(* IEC 61131-3 sources: JingjiangArm/moonboxpro_arm_8.4/Application/Application/任务列表/ExtTask/动作处理/全自动套印2, 17 files *)

(* ---- EnumAutoMaticRegisterCtlMsg.st ---- *)
(*@CES
Name=EnumAutoMaticRegisterCtlMsg
Type=Gvl
TypeGuid=2db5746d-d284-4425-9f7f-2663a34b0ebc
Guid=e7e8891f-fe97-4a56-9291-de397fe1a69c
HasDeclaration=True
HasImplementation=False
*)
{DECLARATION}
// {attribute 'qualified_only'}
// {attribute 'strict'}
TYPE EnumAutoMaticRegisterCtlMsg :
(
	AMRC_MSG_NORMAL := 0,                (* 正常 *)
    AMRC_MSG_ERR_BUSY_HOR,               (* 横向正忙 *)
    AMRC_MSG_ERR_LASTAXISID_INVALID,     (* 最后一个轴id非法 *)
    AMRC_MSG_ERR_AUTOPREGISTER_VER,      (* 自动纵向套印失败 *)
    AMRC_MSG_TIMEOUT_HOR,                (* 横向预套准启动超时状态 *)
    AMRC_MSG_TIMEOUT_WAITPOS_3RD,        (* 第三方设备位置等待超时 *)
    AMRC_MSG_TIMEOUT_WAITPOS_MANU        (* 手动位置等待超时 *)
);
END_TYPE

{IMPLEMENTATION}

(* ---- EnumAutoPrintMasterStep.st ---- *)
(*@CES
Name=EnumAutoPrintMasterStep
Type=Gvl
TypeGuid=2db5746d-d284-4425-9f7f-2663a34b0ebc
Guid=e561adc0-0517-4418-b830-643ab1aeef13
HasDeclaration=True
HasImplementation=False
*)
{DECLARATION}
// 主控制状态机枚举
TYPE EnumAutoPrintMasterStep :
(
    APM_STEP_IDLE := 0,                  (* 1空闲 *)
    APM_STEP_TIPS,                       (* 2提示 *)
    APM_STEP_TIPS_ALARM,                 (* 3警铃提示 *)
    APM_STEP_AUTO_HOR,                   (* 4横向预对版 *)
    APM_STEP_AUTOING_HOR,                (* 5横向对版中 *)
    APM_STEP_AUTOSENSORPOS,              (* 6自动传感器位置 *)
    APM_STEP_SENSORPOSBYSYS3RD,          (* 7第三方设备获取传感器位置 *)
    APM_STEP_WAITPOSBY3RD,               (* 8等待第三方位置 *)
    APM_STEP_SENSORPOSBYMANU,            (* 9手动获取传感器位置 *)
    APM_STEP_WAITPOSBYMANU,              (* 10等待手动位置 *)
    APM_STEP_SENSOR_TO_TARGETPOS,        (* 11传感器到目标位置 *)
    APM_STEP_SENSOR_TO_TARGETPOSING,     (* 12传感器到目标位置中 *)
    APM_STEP_AUTO_VER,                   (* 13纵向全自动套印 *)
    APM_STEP_AUTOING_VER,                (* 14纵向全自动套印中 *)
    APM_STEP_AUTODNE_VER,                (* 15纵向全自动套印完成 *)
	APM_STEP_CALC_ADJUSTMENTS,             (** 16计算调整量 *)
    APM_STEP_FAST_ADJUSTMENT,              (** 17快速对版调整 *)
    APM_STEP_COMPLETE,                     (** 18完成 *)
    APM_STEP_TIMEOUT,                    (* 19超时 *)
    APM_STEP_ERR                         (* 20错误 *)
);
END_TYPE

{IMPLEMENTATION}

(* ---- EnumFindCommand.st ---- *)
(*@CES
Name=EnumFindCommand
Type=Gvl
TypeGuid=2db5746d-d284-4425-9f7f-2663a34b0ebc
Guid=4d4922df-cbf7-48ea-9894-b69efa7c7e4f
HasDeclaration=True
HasImplementation=False
*)
{DECLARATION}
// {attribute 'qualified_only'}
// {attribute 'strict'}
TYPE EnumFindCommand :
(
    FIND_CMD_IDLE := 0,                    (* 空闲 *)
    FIND_CMD_START_SINGLE,                 (* 开始单色寻找 *)
    FIND_CMD_START_MIX,                    (* 开始混色寻找 *)
    FIND_CMD_RESET                         (* 重置 *)
);
END_TYPE
{IMPLEMENTATION}

(* ---- EnumFindErrorCode.st ---- *)
(*@CES
Name=EnumFindErrorCode
Type=Gvl
TypeGuid=2db5746d-d284-4425-9f7f-2663a34b0ebc
Guid=764d2f18-3722-49fd-bd0f-02e1ffafaf8d
HasDeclaration=True
HasImplementation=False
*)
{DECLARATION}
// 寻找错误代码枚举
TYPE EnumFindErrorCode :
(
   	FIND_ERR_NONE := 0,                  (* 无错误 *)
    FIND_ERR_COARSE_NOT_READY := 88,     (* 粗调未到位 *)
    FIND_ERR_WAITING_CIRCLE := 50,       (* 等待1.5圈中 *)
    FIND_ERR_WAITING_FIBER_IDLE := 51,   (* 等待光纤空闲 *)
    FIND_ERR_SINGLE_MARK_NOT_FOUND := 101,(* 单色标记未找到 *)
    FIND_ERR_CALC_BEST_FAILED := 102,    (* 最佳位置计算失败 *)
    FIND_ERR_PRE_POS_INVALID := 103,     (* 前色位置无效 *)
    FIND_ERR_WAITING_SINGLE_INFO := 53,  (* 等待单色新的一圈信息 *)
    FIND_ERR_WAITING_MIX_INFO := 54,     (* 等待前色信息 *)
    FIND_ERR_TIMEOUT := 200,             (* 超时 *)
    FIND_ERR_AXIS_ID_INVALID := 201,     (* 轴ID无效 *)
    FIND_ERR_NOT_ENABLED := 202,         (* 未使能 *)
    FIND_ERR_UNKNOWN := 255              (* 未知错误 *)
);
END_TYPE
{IMPLEMENTATION}

(* ---- EnumFindState.st ---- *)
(*@CES
Name=EnumFindState
Type=Gvl
TypeGuid=2db5746d-d284-4425-9f7f-2663a34b0ebc
Guid=4b638ac6-7ee9-4b1b-9b99-b2600605b011
HasDeclaration=True
HasImplementation=False
*)
{DECLARATION}
// {attribute 'qualified_only'}
// {attribute 'strict'}
// 寻找模块状态
TYPE EnumFindState :
(
    FIND_STATE_IDLE := 0,                (* 0空闲 *)
    FIND_STATE_INIT,                     (* 1初始化 *)
    FIND_STATE_WAIT_PRESS,               (* 2等待合压 *)
    FIND_STATE_CHECK_COARSE,             (* 3检查粗调 *)
    FIND_STATE_DELAY_SINGLE,             (* 4单色前延时 *)
    FIND_STATE_FIND_SINGLE,              (* 5寻找单色 *)
    FIND_STATE_MOVE_FIBER,               (* 6移动光纤 *)
    FIND_STATE_WAIT_FIBER_MOVE,          (* 7等待光纤移动 *)
    FIND_STATE_CALC_BEST,                (* 8计算最佳位置 *)
    FIND_STATE_ADJUST_GATE,              (* 9调整波门 *)
    FIND_STATE_DELAY_MIX,                (* 10混色前延时 *)
    FIND_STATE_FINE_ADJUST,              (* 11光纤精调 *)
    FIND_STATE_WAIT_FINE_ADJ,            (* 12等待精调完成 *)
    FIND_STATE_FIND_MIX,                 (* 13寻找混色 *)
    FIND_STATE_COMPLETE,                 (* 14完成 *)
    FIND_STATE_ERROR                     (* 15错误 *)
);
END_TYPE
{IMPLEMENTATION}

(* ---- StFindResult.st ---- *)
(*@CES
Name=StFindResult
Type=Gvl
TypeGuid=2db5746d-d284-4425-9f7f-2663a34b0ebc
Guid=f624abef-a881-46ee-91b9-f19468406fe9
HasDeclaration=True
HasImplementation=False
*)
{DECLARATION}
{attribute 'pack_mode' := '1'}
// 寻找模块结果
TYPE StFindResult :
STRUCT
    xSuccess: BOOL;                      (* 寻找成功 *)
    iCurLabelPos: INT;                   (* 当前色位置 *)
    iPreLabelPos: INT;                   (* 前色位置 *)
    iCurBestPos: INT;                    (* 当前色最佳位置 *)
    rFiberMoveDist: REAL;                (* 光纤移动距离 *)
    iErrorCode: INT;                     (* 错误代码 *)
	eState: EnumFindState;				(*轴状态*)
    //sErrorMessage: STRING(255);          (* 错误信息 *)
END_STRUCT
END_TYPE
{IMPLEMENTATION}

(* ---- KS_CalBestFiberMoveDisByPS.st ---- *)
(*@CES
Name=KS_CalBestFiberMoveDisByPS
Type=FunctionBlock
TypeGuid=6f9dac99-8de1-4efc-8465-68ac443b7d08
Guid=54f61bec-2d54-4cc2-8835-56cc55fddebe
HasDeclaration=True
HasImplementation=True
*)
{DECLARATION}
FUNCTION KS_CalBestFiberMoveDisByPS : REAL
VAR_INPUT
	i_rwidth      		:POINTER TO REAL;    (*色标宽度*)
	rmark_width      : BYTE;                 (*三角形标宽度*)
    rmark_height     : BYTE;                 (*三角形标高度*)
	i_iMarkId        : INT; (*三角形标类型*)
	i_pBestMoveDisPS: POINTER TO REAL;
END_VAR
VAR
	rstandard_value  : REAL;                 (*标准宽度*)
	rdiff            : REAL;                 (*差值*)
    rdeviation       : REAL;                 (*差值乘比例*)
	rratio           : REAL;                 (*宽高比例*)
	rmove            : REAL;

END_VAR

{IMPLEMENTATION}
// 1. 安全检查：避免除零
IF (rmark_height < 1) THEN
    i_pBestMoveDisPS^ := REAL#-0.0;
    RETURN;
END_IF;

// 1. 安全检查：避免除零
IF (i_rwidth^ = 0) THEN
    i_pBestMoveDisPS^ := REAL#-0.0;
    RETURN;
END_IF;

rstandard_value := BYTE_TO_REAL(rmark_height) / 2.0;
rdiff := i_rwidth^ - rstandard_value;
rratio := BYTE_TO_REAL(rmark_width) / BYTE_TO_REAL(rmark_height);
rmove := rdiff * rratio;

// 4. 根据MARK类型决定方向
IF i_iMarkId = MARK_TYPE_TRAPE_VFLN OR i_iMarkId = MARK_TPYE_TRAPE_VBLN THEN
    i_pBestMoveDisPS^ := -rmove;  // 宽了向左调
ELSIF i_iMarkId = MARK_TYPE_TRAPE_VFLP OR i_iMarkId = MARK_TYPE_TRAPE_VBLP THEN
    i_pBestMoveDisPS^ := rmove;   // 窄了向右调
ELSIF i_iMarkId = MARK_TYPE_LINE THEN (*条标*)
	i_pBestMoveDisPS^ := 0;
END_IF;

(* ---- KS_CalBestFiberMoveDisByRS.st ---- *)
(*@CES
Name=KS_CalBestFiberMoveDisByRS
Type=FunctionBlock
TypeGuid=6f9dac99-8de1-4efc-8465-68ac443b7d08
Guid=ef5f33da-28ef-4533-8c0f-8778b1cdea74
HasDeclaration=True
HasImplementation=True
*)
{DECLARATION}
FUNCTION KS_CalBestFiberMoveDisByRS : REAL
VAR_INPUT
	i_ar_width       : ARRAY[1..3] OF REAL;    (*三个位置的色标宽度*)
	i_ar_markerpos   : ARRAY[1..3] OF INT;     (*三个色标位置信息*)
	rmark_width      : BYTE;                 (*三角形标宽度*)
    rmark_height     : BYTE;                 (*三角形标高度*)
	i_iMarkId        : INT; (*三角形标类型*)
	i_pBestPositionRS : POINTER TO INT;
	i_pBestMoveDisRS: POINTER TO REAL;
END_VAR
VAR
	i_ar_position : ARRAY[1..3] OF REAL := [0.0,-3.0,3.0];
	rstandard_value  : REAL;                 (*标准宽度*)
    ibest_index      : INT := -1;            // 最佳点索引
    rmin_diff        : REAL := REAL#1.0E6;   // 最小差值（初始值）
    iN              : INT;                   // 循环计数器
    rcurrent_diff    : REAL;                  // 当前循环计算的差值
    rbest_width      : REAL;                  // 最佳点对应的宽度
    rbest_pos        : REAL;                  // 最佳点对应的位置
    rcurrent_pos     : REAL;                  // 当前机械位置
    rwidth_ratio     : REAL;                  // 宽高比
    rdeviation       : REAL;                  // 计算出的偏差量
    rtarget_pos      : REAL;                  // 最终目标位置

END_VAR

{IMPLEMENTATION}
// 1. 安全检查：避免除零
IF (rmark_height < 1) THEN
    i_pBestMoveDisRS^ := REAL#-3.0;
    RETURN;
END_IF;

// 2. 遍历筛选最佳点（宽度最接近标准值）
ibest_index := -1;
rmin_diff := REAL#1.0E6;
rstandard_value := BYTE_TO_REAL(rmark_height) / 2;

FOR iN := 1 TO 3 DO
    // 假设位置为 -1.0 或者宽度为 -0.0 表示该点无效
    IF (i_ar_markerpos[iN] = -1 OR i_ar_width[iN] = REAL#0.0) THEN
		CONTINUE;
	ELSE
        rcurrent_diff := ABS(i_ar_width[iN] - rstandard_value);
        // 更新最佳点
        IF (rcurrent_diff < rmin_diff) THEN
            rmin_diff := rcurrent_diff;
            ibest_index := iN;
        END_IF;
    END_IF;
END_FOR;

// 3. 若无有效点，退回原点
IF (ibest_index < 0) THEN
    i_pBestMoveDisRS^ := REAL#-3.0;
    RETURN;
END_IF;

// 4. 提取计算所需数据
rbest_width := i_ar_width[ibest_index];
rbest_pos := i_ar_position[ibest_index];
rcurrent_pos := i_ar_position[3]; // 当前位置锁定为第三个点 (Index 2)

// 5. 计算几何偏差
rwidth_ratio := BYTE_TO_REAL(rmark_width) / BYTE_TO_REAL(rmark_height);
rdeviation := rmin_diff * rwidth_ratio;

// 6. 确定目标位置   以后可以改成根据色标形式控制左右方向   总体而言，是宽了往窄的方向移动，窄了往宽的方向移动
IF (i_iMarkId = MARK_TYPE_TRAPE_VFLN OR i_iMarkId = MARK_TPYE_TRAPE_VBLN) THEN
	IF (rbest_width > rstandard_value) THEN
		rtarget_pos := rbest_pos - rdeviation; // 太宽 -> 向左
	ELSIF (rbest_width < rstandard_value) THEN
		rtarget_pos := rbest_pos + rdeviation; // 太窄 -> 向右
	ELSE
		rtarget_pos := rbest_pos; // 正好
	END_IF;
ELSIF (i_iMarkId = MARK_TYPE_TRAPE_VFLP OR i_iMarkId = MARK_TYPE_TRAPE_VBLP) THEN
	IF (rbest_width > rstandard_value) THEN
		rtarget_pos := rbest_pos + rdeviation; // 太宽 -> 向右
	ELSIF (rbest_width < rstandard_value) THEN
		rtarget_pos := rbest_pos - rdeviation; // 太窄 -> 向左
	ELSE
		rtarget_pos := rbest_pos; // 正好
	END_IF;
ELSIF i_iMarkId = MARK_TYPE_LINE THEN (*条标*)
	FOR iN := 1 TO 3 DO
		// 假设位置为 -1.0 或者宽度为 -1.0 表示该点无效
		IF (i_ar_markerpos[iN] = -1 OR i_ar_width[iN] = REAL#-1.0) THEN
			CONTINUE;
		ELSE
			ibest_index := iN;
			EXIT;
		END_IF;
	END_FOR;
	(*这样可以回到零位*)
	rtarget_pos:= 0;
END_IF

// 7. 计算并返回最终移动距离
i_pBestMoveDisRS^ := rtarget_pos - rcurrent_pos;
i_pBestPositionRS^ := i_ar_markerpos[ibest_index];

(* ---- KS_CalculateMixFindDelayTime.st ---- *)
(*@CES
Name=KS_CalculateMixFindDelayTime
Type=FunctionBlock
TypeGuid=6f9dac99-8de1-4efc-8465-68ac443b7d08
Guid=2d7bebb1-5781-4f9d-9266-922f12b4caec
HasDeclaration=True
HasImplementation=True
*)
{DECLARATION}
FUNCTION KS_CalculateMixFindDelayTime  : uint
VAR_INPUT
    i_iAxisId: INT;                        (* 轴号 *)
    i_iBeforeAxisId: INT;                  (* 前轴号 *)
    i_pstUnitParam_Save: POINTER TO StUnitParam_Save; (* 单元参数 *)
    i_rVel: REAL;                          (* 速度 *)
END_VAR
VAR
    uiDelayTime: UINT;                     (* 延时时间@ms *)
    pstUnitParam_Save: POINTER TO StUnitParam_Save;
    rWaitTime: REAL;                       (* 等待时间@s *)
    rFilmLength: REAL;                     (* 料长@m *)
END_VAR
{IMPLEMENTATION}
pstUnitParam_Save := i_pstUnitParam_Save;
uiDelayTime := 0;

(* 计算前一色到此色的料长 *)
IF i_iBeforeAxisId <> -1 THEN
    (* 获取前一色到此色的料长 *)
    rFilmLength := (pstUnitParam_Save^.rFilmLengthFromPrevPressUnit)/1000.0*(i_iAxisId-i_iBeforeAxisId);

    (* 计算等待时间：料长(m) / 速度(m/min) * 60s/min = 等待时间(s) *)
    IF i_rVel > 0 THEN
        rWaitTime := rFilmLength / i_rVel * 60.0;

        (* 转换为毫秒 *)
        uiDelayTime := REAL_TO_UINT(rWaitTime * 1000.0);
    ELSE
        (* 速度为零，使用默认值 *)
        uiDelayTime := 30000;  (* 30秒 *)
    END_IF
END_IF

(* 增加安全余量（5个版周长的时间） *)
IF pstUnitParam_Save^.rGirth_PrnRoller > 0 AND i_rVel > 0 THEN
    rWaitTime := 5.0 * pstUnitParam_Save^.rGirth_PrnRoller / 1000.0 / i_rVel * 60.0;
    uiDelayTime := uiDelayTime + REAL_TO_UINT(rWaitTime * 1000.0);
END_IF

(* 最小延时时间 *)
IF uiDelayTime < 1000 THEN
    uiDelayTime := 1000;  (* 至少1秒 *)
END_IF

KS_CalculateMixFindDelayTime := uiDelayTime;

(* ---- KS_CalculateVerticalAdjustment.st ---- *)
(*@CES
Name=KS_CalculateVerticalAdjustment
Type=FunctionBlock
TypeGuid=6f9dac99-8de1-4efc-8465-68ac443b7d08
Guid=55283c42-1c2e-4d65-8dd3-8f793fe68a41
HasDeclaration=True
HasImplementation=True
*)
{DECLARATION}
(*返回计算误差的点数*)
FUNCTION KS_CalculateVerticalAdjustment : real
VAR_INPUT
    i_iAxisId: INT;                        (* 轴号 *)
    i_iCurBestSignalPos: INT;              (* 当前色最佳位置 *)
    i_iPreLabelPos: INT;                   (* 前色位置 *)
    i_pstUnitParam_Save: POINTER TO StUnitParam_Save; (* 单元参数 *)
    i_pstGrpParam_Save: POINTER TO StGrpParam_Save;  (* 组参数 *)
END_VAR
VAR
   	rAdjValue: REAL;                       (* 调整量@粗采样点数*)
    pstUnitParam_Save: POINTER TO StUnitParam_Save;
    pstGrpParam_Save: POINTER TO StGrpParam_Save;
    rTmp: REAL;
END_VAR
{IMPLEMENTATION}
pstUnitParam_Save := i_pstUnitParam_Save;
pstGrpParam_Save := i_pstGrpParam_Save;

(* 初始化返回值 *)
rAdjValue := 0.0;

(* 检查输入有效性 *)
IF i_iCurBestSignalPos >= 0 AND i_iPreLabelPos >= 0 AND
   i_iCurBestSignalPos < 4000 AND i_iPreLabelPos < 4000 THEN

    (* 根据标记排列方式计算调整量 *)
    IF pstUnitParam_Save^.iMarkArrangeMode = MARK_ARRANGE_VFOR THEN
        (* 正向排列 *)
        rTmp := INT_TO_REAL(i_iCurBestSignalPos - i_iPreLabelPos -
                   LREAL_TO_INT(20.0 * MAX_ROUNDSAMPLE_NUM / pstUnitParam_Save^.rGirth_PrnRoller));
    ELSIF pstUnitParam_Save^.iMarkArrangeMode = MARK_ARRANGE_VREV THEN
        (* 反向排列 *)
        rTmp := INT_TO_REAL(i_iCurBestSignalPos - i_iPreLabelPos +
                   LREAL_TO_INT(20.0 * MAX_ROUNDSAMPLE_NUM / pstUnitParam_Save^.rGirth_PrnRoller));
    ELSE
        (* 默认处理 *)
        rTmp := INT_TO_REAL(i_iCurBestSignalPos - i_iPreLabelPos);
    END_IF

    (* 将调整的粗采样点数转换到±MAX_ROUNDSAMPLE_NUM/2范围内 *)
    WHILE rTmp < -MAX_ROUNDSAMPLE_NUM / 2.0 DO
        rTmp := rTmp + MAX_ROUNDSAMPLE_NUM;
    END_WHILE
    WHILE rTmp > MAX_ROUNDSAMPLE_NUM / 2.0 DO
        rTmp := rTmp - MAX_ROUNDSAMPLE_NUM;
    END_WHILE

    (* 计算um单位：调整量(um) = 点数 * 版辊周长(um) / 总采样点数 *)
   // rAdjValue := rTmp * pstUnitParam_Save^.rGirth_PrnRoller * 1000.0 / MAX_ROUNDSAMPLE_NUM;
END_IF

KS_CalculateVerticalAdjustment := rTmp;

(* ---- KS_CheckSensorMotorIdleSts.st ---- *)
(*@CES
Name=KS_CheckSensorMotorIdleSts
Type=FunctionBlock
TypeGuid=6f9dac99-8de1-4efc-8465-68ac443b7d08
Guid=e3f21590-970b-415a-a0bb-786d7afe314f
HasDeclaration=True
HasImplementation=True
*)
{DECLARATION}
FUNCTION KS_CheckSensorMotorIdleSts : BOOL
(*|=0 检查所有传感器的是否处于空闲状态@所有都空闲则输出true|有一个在运动就置位false*)
(*|=合法轴id,则返回轴状态|TRUE 是空闲,FALSE是运动*)
VAR_INPUT
	i_iAxisId:INT;(*轴号@=0 *)
	i_byAxisNum:BYTE;(*轴个数@全自动套印轴*)
	i_aiAxisList_AutoAdj:ARRAY [1..MAX_UNIT_NUM] OF int;(*轴列表*)
	i_axSensorMotorIdle:ARRAY [1..MAX_UNIT_NUM] OF BOOL;(*传感器电机空闲状态@该状态不是直接通讯上来的,需要做处理后的*)
END_VAR
VAR
	iN: INT;
	xSensorMotorIdle: BOOL;
	iAxisId: INT;
	xResult: BOOL:=TRUE;
END_VAR
{IMPLEMENTATION}
IF i_iAxisId=0 THEN
	FOR iN:=2 TO i_byAxisNum BY 1 DO
		iAxisId:=i_aiAxisList_AutoAdj[iN];
		IF iAxisId>0 AND iAxisId<=MAX_UNIT_NUM THEN
			xSensorMotorIdle:=i_axSensorMotorIdle[iAxisId];
			IF NOT xSensorMotorIdle THEN(*处于运动中*)
				xResult:=FALSE;
				EXIT;
			END_IF
		END_IF
	END_FOR
ELSE
	iAxisId:=i_iAxisId;
	IF iAxisId>0 AND iAxisId<=MAX_UNIT_NUM THEN
		xSensorMotorIdle:=i_axSensorMotorIdle[iAxisId];
		IF NOT xSensorMotorIdle THEN(*处于运动中*)
			xResult:=FALSE;
		END_IF
	END_IF
END_IF

KS_CheckSensorMotorIdleSts:=xResult;

(* ---- KS_CreateTemplate.st ---- *)
(*@CES
Name=KS_CreateTemplate
Type=FunctionBlock
TypeGuid=6f9dac99-8de1-4efc-8465-68ac443b7d08
Guid=90238752-c97b-4d95-b35e-1bfe3f1964c0
HasDeclaration=True
HasImplementation=True
*)
{DECLARATION}
//构建模版函数
FUNCTION KS_CreateTemplate : BOOL
VAR_INPUT
	i_bySignalType : byte;(*模版类型，1 北人标，2普通标 ，3科赛引导条标*)
	i_iMarkTypeId : INT;(*色标形式pstStGrpParam_Save^.iMarkTypeId*)
	i_iMarkArrangeMode :INT;(*顺逆序输入*)
	i_byColorIdCurrent						: BYTE;(*当前轴色序*)
	i_rGirth_PrnRoller        :REAL;(*版周*)
	//模版构建方法 要求条标直接输入起点mm与终点mm，三角标，先确定直角边的位置，斜边按照三角标高度的一半推
	i_paiModeMidPoint:POINTER TO ARRAY [1..4] OF INT;
	i_pabyModeRadius:POINTER TO ARRAY [1..4] OF BYTE;
	i_parModeStartmm: POINTER TO ARRAY [1..4] OF REAL;
	i_parModeEndmm:POINTER TO ARRAY [1..4] OF REAL;
	i_parSignalMsg:POINTER TO ARRAY [1..15] OF REAL;
END_VAR
VAR
	iN:INT;//循环计数
	rMaxEndTemp:REAL;//记录一下最大坐标
	arStart1UMM: ARRAY [1..4] OF REAL; //mm单位 规定顺序 旗标 id 1  圆标 id 2  引导标 id 3  三角标 id 4
	arEnd1UMM: ARRAY [1..4] OF REAL; //mm单位 规定顺序 旗标 id 1  圆标 id 2  引导标 id 3  三角标 id 4
	arStart2UMM: ARRAY [1..4] OF REAL; //mm单位 规定顺序 旗标 id 1  圆标 id 2  引导标 id 3  三角标 id 4
	arEnd2UMM:ARRAY [1..4] OF REAL; //mm单位 规定顺序 旗标 id 1  圆标 id 2  引导标 id 3  三角标 id 4
	arStartMM: ARRAY [1..4] OF REAL; //mm单位 规定顺序 旗标 id 1  圆标 id 2  引导标 id 3  三角标 id 4
	arEndMM: ARRAY [1..4] OF REAL; //mm单位 规定顺序 旗标 id 1  圆标 id 2  引导标 id 3  三角标 id 4
	arStartMMTemp: ARRAY [1..4] OF REAL; //mm单位 用来导逆序，规定顺序 旗标 id 1  圆标 id 2  引导标 id 3  三角标 id 4
	arEndMMTemp: ARRAY [1..4] OF REAL; //mm单位 用来导逆序，规定顺序 旗标 id 1  圆标 id 2  引导标 id 3  三角标 id 4
	arSignalMsg:ARRAY [1..15] OF REAL; (*1旗标高度
										2 圆标高度
										3 2色引导标高度
										4 三角标高度
										5 1色旗标终点-圆标起点
										6 2色旗标终点-圆标起点
										7 1色圆标终点-引导标起点
										8 2色圆标终点-引导标起点
										9 1色引导标终点-三角标起点
										10 2色引导标终点-三角标起点
										11 2色引导标起点点-3色引导标起点
										12 1色引导标高度
*)

END_VAR

{IMPLEMENTATION}

IF 	i_parSignalMsg <> 0 AND i_rGirth_PrnRoller <> 0  THEN
	arSignalMsg:=i_parSignalMsg^;

	CASE i_bySignalType OF
	1:	//科赛引导标
		//先构建1色的模版
		arStart1UMM[1]:=  arSignalMsg[1] /2.0;//旗标起点定义旗标高度一半
		arEnd1UMM[1]:= arSignalMsg[1];//旗标终点定义旗标终点
		arStart1UMM[2]:= arEnd1UMM[1] + arSignalMsg[5];//圆标起点为旗标终点+1u5
		arEnd1UMM[2]:= arStart1UMM[2] + arSignalMsg[2];
		arStart1UMM[3]:= arEnd1UMM[2] + arSignalMsg[7];
		arEnd1UMM[3]:= arStart1UMM[3] + arSignalMsg[12];
		//条标
		IF i_iMarkTypeId = MARK_TYPE_LINE THEN
			arStart1UMM[4]:= arEnd1UMM[3] + arSignalMsg[9];
			arEnd1UMM[4]:= arStart1UMM[4] + arSignalMsg[4];
		//直角边在前
		ELSIF i_iMarkTypeId = MARK_TYPE_TRAPE_VFLP OR  i_iMarkTypeId = MARK_TYPE_TRAPE_VFLN THEN
			arStart1UMM[4]:= arEnd1UMM[3] + arSignalMsg[9];
			arEnd1UMM[4]:= arStart1UMM[4] + arSignalMsg[4]/2.0;
		ELSIF  i_iMarkTypeId = MARK_TYPE_TRAPE_VBLP OR  i_iMarkTypeId = MARK_TPYE_TRAPE_VBLN THEN
		//直角边在后
			arStart1UMM[4]:= arEnd1UMM[3] + arSignalMsg[9]+arSignalMsg[4]/2.0;
			arEnd1UMM[4]:=  arEnd1UMM[3] + arSignalMsg[9]+arSignalMsg[4];
		END_IF
		//构建2色的模版
		arStart2UMM[1]:=  arSignalMsg[1] /2.0;//旗标起点定义旗标高度一半
		arEnd2UMM[1]:= arSignalMsg[1];//旗标终点定义旗标终点
		arStart2UMM[2]:= arEnd2UMM[1] + arSignalMsg[6];
		arEnd2UMM[2]:= arStart2UMM[2] + arSignalMsg[2];
		arStart2UMM[3]:= arEnd2UMM[2] + arSignalMsg[8];
		arEnd2UMM[3]:= arStart2UMM[3] + arSignalMsg[3];
		//条标
		IF i_iMarkTypeId = MARK_TYPE_LINE THEN
			arStart2UMM[4]:= arEnd1UMM[3] + arSignalMsg[10];
			arEnd2UMM[4]:= arEnd1UMM[3] + arSignalMsg[10]+(arSignalMsg[4]);
		ELSIF i_iMarkTypeId = MARK_TYPE_TRAPE_VFLP OR  i_iMarkTypeId = MARK_TYPE_TRAPE_VFLN THEN
			arStart2UMM[4]:= arEnd1UMM[3] + arSignalMsg[10];
			arEnd2UMM[4]:= arEnd1UMM[3] + arSignalMsg[10]+(arSignalMsg[4]/2.0);
		ELSIF i_iMarkTypeId = MARK_TYPE_TRAPE_VBLP OR i_iMarkTypeId = MARK_TPYE_TRAPE_VBLN THEN
		//直角边在后
			arStart2UMM[4]:= arEnd1UMM[3] + arSignalMsg[10]+arSignalMsg[4]/2.0;
			arEnd2UMM[4]:=  arEnd1UMM[3] + arSignalMsg[10]+arSignalMsg[4];
		END_IF
		IF i_byColorIdCurrent > 0 THEN
			//根据色序选择模版
			CASE i_byColorIdCurrent OF
				1:
					FOR iN := 1 TO 4 BY 1 DO
						arStartMM[iN]:=arStart1UMM[iN];
						arEndMM[iN]:=arEnd1UMM[iN];
					END_FOR
				2:
					FOR iN := 1 TO 4 BY 1 DO
						arStartMM[iN]:=arStart2UMM[iN];
						arEndMM[iN]:=arEnd2UMM[iN];
					END_FOR
				ELSE
					arStartMM[1]:=arStart1UMM[1];
					arEndMM[1]:=arEnd1UMM[1];
					arStartMM[2]:=arStart1UMM[2]+(i_byColorIdCurrent-1)*(arSignalMsg[6]-arSignalMsg[5]);
					arEndMM[2]:=arEnd1UMM[2]+(i_byColorIdCurrent-1)*(arSignalMsg[6]-arSignalMsg[5]);
					arStartMM[3]:=arStart1UMM[3]+(i_byColorIdCurrent-1)*(arStart2UMM[3]-arStart1UMM[3]);
					arEndMM[3]:=arEnd1UMM[3]+(i_byColorIdCurrent-1)*(arEnd2UMM[3]-arEnd1UMM[3]);
					arStartMM[4]:=arStart1UMM[4]+(i_byColorIdCurrent-1)*(arStart2UMM[4]-arStart1UMM[4]);
					arEndMM[4]:=arEnd1UMM[4]+(i_byColorIdCurrent-1)*(arEnd2UMM[4]-arEnd1UMM[4]);
			END_CASE
		ELSE
			FOR iN := 1 TO 4 BY 1 DO
				arStartMM[iN]:=0;
				arEndMM[iN]:=0;
			END_FOR
		END_IF
	2: //普通标
		//关于建立没有引导,只有旗标，圆标，三角标，标建立模版，要求 3,7,8,11,12均为0，9,10填写圆标到三角标的距离，模版建立方法，虚拟一个引导标，将引导标的起点和终点与三角标相同
		//先构建1色的模版
		arStart1UMM[1]:=  arSignalMsg[1] /2.0;//旗标起点定义旗标高度一半
		arEnd1UMM[1]:= arSignalMsg[1];//旗标终点定义旗标终点
		arStart1UMM[2]:= arEnd1UMM[1] + arSignalMsg[5];//圆标起点为旗标终点+1u5
		arEnd1UMM[2]:= arStart1UMM[2] + arSignalMsg[2];

		//条标
		IF i_iMarkTypeId = MARK_TYPE_LINE THEN
			arStart1UMM[4]:= arEnd1UMM[2] + arSignalMsg[9];
			arEnd1UMM[4]:= arStart1UMM[4] + arSignalMsg[4];
			arStart1UMM[3]:= arStart1UMM[4];
			arEnd1UMM[3]:= arEnd1UMM[4];
		//直角边在前
		ELSIF i_iMarkTypeId = MARK_TYPE_TRAPE_VFLP OR  i_iMarkTypeId = MARK_TYPE_TRAPE_VFLN THEN
			arStart1UMM[4]:= arEnd1UMM[2] + arSignalMsg[9];
			arEnd1UMM[4]:= arStart1UMM[4] + arSignalMsg[4]/2.0;
			arStart1UMM[3]:= arStart1UMM[4];
			arEnd1UMM[3]:= arEnd1UMM[4];
		ELSIF  i_iMarkTypeId = MARK_TYPE_TRAPE_VBLP OR  i_iMarkTypeId = MARK_TPYE_TRAPE_VBLN THEN
		//直角边在后
			arStart1UMM[4]:= arEnd1UMM[2] + arSignalMsg[9]+arSignalMsg[4]/2.0;
			arEnd1UMM[4]:=  arEnd1UMM[2] + arSignalMsg[9]+arSignalMsg[4];
			arStart1UMM[3]:= arStart1UMM[4];
			arEnd1UMM[3]:= arEnd1UMM[4];
		END_IF
		//构建2色的模版
		arStart2UMM[1]:=  arSignalMsg[1] /2.0;//旗标起点定义旗标高度一半
		arEnd2UMM[1]:= arSignalMsg[1];//旗标终点定义旗标终点
		arStart2UMM[2]:= arEnd2UMM[1] + arSignalMsg[6];
		arEnd2UMM[2]:= arStart2UMM[2] + arSignalMsg[2];
		//条标
		IF i_iMarkTypeId = MARK_TYPE_LINE THEN
			arStart2UMM[4]:= arEnd2UMM[2] + arSignalMsg[10];
			arEnd2UMM[4]:= arStart2UMM[4] + arSignalMsg[4];
			arStart2UMM[3]:=arStart2UMM[4];
			arEnd2UMM[3]:= arEnd2UMM[4];
		//直角边在前
		ELSIF i_iMarkTypeId = MARK_TYPE_TRAPE_VFLP OR  i_iMarkTypeId = MARK_TYPE_TRAPE_VFLN THEN
			arStart2UMM[4]:= arEnd2UMM[2] + arSignalMsg[10];
			arEnd2UMM[4]:= arStart2UMM[4] + arSignalMsg[4]/2.0;
			arStart2UMM[3]:=arStart2UMM[4];
			arEnd2UMM[3]:= arEnd2UMM[4];
		ELSIF i_iMarkTypeId = MARK_TYPE_TRAPE_VBLP OR i_iMarkTypeId = MARK_TPYE_TRAPE_VBLN THEN
		//直角边在后
			arStart2UMM[4]:= arEnd2UMM[2] + arSignalMsg[10]+arSignalMsg[4]/2.0;
			arEnd2UMM[4]:=  arEnd2UMM[2] + arSignalMsg[10]+arSignalMsg[4];
			arStart2UMM[3]:=arStart2UMM[4];
			arEnd2UMM[3]:= arEnd2UMM[4];
		END_IF
		IF i_byColorIdCurrent > 0 THEN
			//根据色序选择模版
			CASE i_byColorIdCurrent OF
				1:
					FOR iN := 1 TO 4 BY 1 DO
						arStartMM[iN]:=arStart1UMM[iN];
						arEndMM[iN]:=arEnd1UMM[iN];
					END_FOR
				2:
					FOR iN := 1 TO 4 BY 1 DO
						arStartMM[iN]:=arStart2UMM[iN];
						arEndMM[iN]:=arEnd2UMM[iN];
					END_FOR
				ELSE
					arStartMM[1]:=arStart1UMM[1];
					arEndMM[1]:=arEnd1UMM[1];
					arStartMM[2]:=arStart1UMM[2]+(i_byColorIdCurrent-1)*(arSignalMsg[6]-arSignalMsg[5]);
					arEndMM[2]:=arEnd1UMM[2]+(i_byColorIdCurrent-1)*(arSignalMsg[6]-arSignalMsg[5]);
					arStartMM[4]:=arStart1UMM[4]+(i_byColorIdCurrent-1)*(arStart2UMM[4]-arStart1UMM[4]);
					arEndMM[4]:=arEnd1UMM[4]+(i_byColorIdCurrent-1)*(arEnd2UMM[4]-arEnd1UMM[4]);
					arStartMM[3]:= arStartMM[4];
					arEndMM[3]:= arEndMM[4];
			END_CASE
		ELSE
			FOR iN := 1 TO 4 BY 1 DO
				arStartMM[iN]:=0;
				arEndMM[iN]:=0;
			END_FOR
		END_IF
	3: // 3 北人标
		//先构建1色的模版
		arStart1UMM[1]:=  arSignalMsg[1] /2.0;//旗标起点定义旗标高度一半
		arEnd1UMM[1]:= arSignalMsg[1];//旗标终点定义旗标终点
		arStart1UMM[2]:= arEnd1UMM[1] + arSignalMsg[5];//圆标起点为旗标终点+1u5
		arEnd1UMM[2]:= arStart1UMM[2] + arSignalMsg[2];
		arStart1UMM[3]:= arEnd1UMM[2] + arSignalMsg[7];
		arEnd1UMM[3]:= arStart1UMM[3] + arSignalMsg[12];
		//条标
		IF i_iMarkTypeId = MARK_TYPE_LINE THEN
			arStart1UMM[4]:= arEnd1UMM[3] + arSignalMsg[9];
			arEnd1UMM[4]:= arStart1UMM[4] + arSignalMsg[4];
		//直角边在前
		ELSIF i_iMarkTypeId = MARK_TYPE_TRAPE_VFLP OR  i_iMarkTypeId = MARK_TYPE_TRAPE_VFLN THEN
			arStart1UMM[4]:= arEnd1UMM[3] + arSignalMsg[9];
			arEnd1UMM[4]:= arStart1UMM[4] + arSignalMsg[4]/2.0;
		ELSIF  i_iMarkTypeId = MARK_TYPE_TRAPE_VBLP OR  i_iMarkTypeId = MARK_TPYE_TRAPE_VBLN THEN
		//直角边在后
			arStart1UMM[4]:= arEnd1UMM[3] + arSignalMsg[9]+arSignalMsg[4]/2.0;
			arEnd1UMM[4]:=  arEnd1UMM[3] + arSignalMsg[9]+arSignalMsg[4];
		END_IF
		//构建2色的模版
		arStart2UMM[1]:=  arSignalMsg[1] /2.0;//旗标起点定义旗标高度一半
		arEnd2UMM[1]:= arSignalMsg[1];//旗标终点定义旗标终点
		arStart2UMM[2]:= arEnd2UMM[1] + arSignalMsg[6];
		arEnd2UMM[2]:= arStart2UMM[2] + arSignalMsg[2];
		arStart2UMM[3]:= arEnd2UMM[2] + arSignalMsg[8];
		arEnd2UMM[3]:= arStart2UMM[3] + arSignalMsg[3];
		//条标
		IF i_iMarkTypeId = MARK_TYPE_LINE THEN
			arStart2UMM[4]:= arEnd1UMM[3] + arSignalMsg[10];
			arEnd2UMM[4]:= arStart1UMM[4] + arSignalMsg[4];
		//直角边在前
		ELSIF i_iMarkTypeId = MARK_TYPE_TRAPE_VFLP OR  i_iMarkTypeId = MARK_TYPE_TRAPE_VFLN THEN
			arStart2UMM[4]:= arEnd2UMM[3] + arSignalMsg[10];
			arEnd2UMM[4]:= arStart2UMM[4] + arSignalMsg[4]/2.0;
		ELSIF i_iMarkTypeId = MARK_TYPE_TRAPE_VBLP OR i_iMarkTypeId = MARK_TPYE_TRAPE_VBLN THEN
		//直角边在后
			arStart2UMM[4]:= arEnd1UMM[3] + arSignalMsg[10]+arSignalMsg[4]/2.0;
			arEnd2UMM[4]:=  arEnd1UMM[3] + arSignalMsg[10]+arSignalMsg[4];
		END_IF
		IF i_byColorIdCurrent > 0 THEN
			//根据色序选择模版
			CASE i_byColorIdCurrent OF
				1:
					FOR iN := 1 TO 4 BY 1 DO
						arStartMM[iN]:=arStart1UMM[iN];
						arEndMM[iN]:=arEnd1UMM[iN];
					END_FOR
				2:
					FOR iN := 1 TO 4 BY 1 DO
						arStartMM[iN]:=arStart2UMM[iN];
						arEndMM[iN]:=arEnd2UMM[iN];
					END_FOR
				ELSE
					arStartMM[1]:=arStart1UMM[1];
					arEndMM[1]:=arEnd1UMM[1];
					arStartMM[2]:=arStart1UMM[2]+(i_byColorIdCurrent-1)*(arSignalMsg[6]-arSignalMsg[5]);
					arEndMM[2]:=arEnd1UMM[2]+(i_byColorIdCurrent-1)*(arSignalMsg[6]-arSignalMsg[5]);
					arStartMM[3]:=arStart2UMM[3]-(i_byColorIdCurrent-2)*arSignalMsg[11];
					arEndMM[3]:=arEnd2UMM[3]-(i_byColorIdCurrent-2)*arSignalMsg[11];
					arStartMM[4]:=arStart2UMM[4]+(i_byColorIdCurrent-2)*(arStart2UMM[4]-arStart1UMM[4]);
					arEndMM[4]:=arEnd2UMM[4]+(i_byColorIdCurrent-2)*(arEnd2UMM[4]-arEnd1UMM[4]);
			END_CASE
		ELSE
			FOR iN := 1 TO 4 BY 1 DO
				arStartMM[iN]:=0;
				arEndMM[iN]:=0;
			END_FOR
		END_IF
	END_CASE
	//根据顺序生成逆序模版
	IF i_iMarkArrangeMode = MARK_ARRANGE_VFOR THEN
		;//不做处理，因为本身构建是顺序的
	ELSIF i_iMarkArrangeMode = MARK_ARRANGE_VREV THEN
		FOR iN := 1 TO 4 BY 1 DO //先记录一下顺序模版
			arStartMMTemp[iN]:=arStartMM[iN];
			arEndMMTemp[iN]:=arEndMM[iN];
		END_FOR
		rMaxEndTemp:= arEndMM[4];
		FOR iN := 1 TO 4 BY 1 DO //导出逆序
			arStartMM[iN]:=rMaxEndTemp-arEndMMTemp[4-iN+1];
			arEndMM[iN]:=rMaxEndTemp-arStartMMTemp[4-iN+1];
		END_FOR
	END_IF
	FOR iN := 1 TO 4 BY 1 DO  //传出中心半径
		i_paiModeMidPoint^[iN]:=REAL_TO_INT((arEndMM[iN]+arStartMM[iN])/2.0/i_rGirth_PrnRoller*MAX_ROUNDSAMPLE_NUM);
		i_pabyModeRadius^[iN]:=REAL_TO_BYTE((arEndMM[iN]-arStartMM[iN])/2.0/i_rGirth_PrnRoller*MAX_ROUNDSAMPLE_NUM);
	END_FOR
	i_parModeStartmm^:=	arStartMM;
	i_parModeEndmm^:=arEndMM;
END_IF

(* ---- KS_FB_AutoPrintMaster.st ---- *)
(*@CES
Name=KS_FB_AutoPrintMaster
Type=FunctionBlock
TypeGuid=6f9dac99-8de1-4efc-8465-68ac443b7d08
Guid=8faa04dc-26bf-43df-9e4a-ef930424aed8
HasDeclaration=True
HasImplementation=True
*)
{DECLARATION}
FUNCTION_BLOCK KS_FB_AutoPrintMaster
VAR_INPUT
    (* 基本输入 *)
    i_xEn: BOOL;                         (* 主使能 *)
    i_rVel: REAL;                        (* 料膜速度@m/min *)
    i_rMachineryFilmLenth: REAL;         (* 机器总料长@m *)
    i_xTipsConfirm: BOOL;                (* 提示确认标志@沿触发 *)
    i_xUseAutoPreRegister_Hor: BOOL;     (* 使用横向对版功能 *)
    i_xAutoPreRegisterIdle_Hor: BOOL;    (* 横向预对版空闲状态 *)
    i_xAutoPreRegistering_Hor: BOOL;     (* 横向预对版中 *)
    i_xUseAutoSensorPos: BOOL;           (* 自动传感器位置@否则直接到纵向全自动纵向套印 *)
    i_xUseSensorPos_3rd: BOOL;           (* 使用第三方设备位置@在线|否则手动移动 *)
    i_xSensorPosValid_3rd: BOOL;         (* 传感器位置有效 *)
    i_rSenserPos_3rd: REAL;              (* 传感器位置@单位未知,暂定一个值 *)
    i_xSensorPosValid_Manu: BOOL;        (* 手动传感器值有效 *)
    i_rSensorPos_Manu: REAL;             (* 手动传感器值@绝对位置@mm *)
    i_xUseFindBestPosStep: BOOL;         (* 使用寻找最佳位置步 *)
	i_xSwitch_RFailure: BOOL;            (** R失效开关 **)
    i_xSwitch_FFailure: BOOL;            (** F失效开关 **)

    (* 轴配置 *)
    i_byAxisNum: BYTE;                   (* 轴个数@全自动套印轴 *)
    i_aiAxisList: ARRAY [1..MAX_UNIT_NUM] OF INT; (* 轴列表 *)
    i_pafbKS_FB_AxisFindModule: POINTER TO ARRAY[1..MAX_UNIT_NUM] OF KS_FB_AxisFindModule;

    (* 系统参数 *)
    i_pstStSysParam: POINTER TO StSysParam;
    i_pastStIOMap_AxisBasic: POINTER TO ARRAY [1..MAX_UNIT_NUM] OF StIOMap_Axis_FE;

    (* 快速对版参数 *)
    i_pastStAxisRapidAdjProf_V: POINTER TO ARRAY[1..MAX_UNIT_NUM] OF StAxisRapidAdjProf_V; (* 快速对版参数数组 *)

    (* 轴状态输入 *)
    i_abyRapidAdjustStep: ARRAY[1..MAX_UNIT_NUM] OF BYTE; (* 各轴快速对版步骤 *)
	i_pastFindResults :POINTER TO ARRAY[1..MAX_UNIT_NUM] OF StFindResult;
END_VAR
VAR_OUTPUT
    (* 状态输出 *)
    o_xEning: BOOL;                      (* 使能中 *)
    o_xAlarm: BOOL;                      (* 3s响铃输出 *)
   // o_xWaitingFilmLenthEn: BOOL;         (* 等料长使能 *)
    o_xAutoPreRegister_Hor: BOOL;        (* 横向自动对版@启动预套后复位 *)
   // o_xExcuteRollerPress_LastAxis: BOOL; (* 最后一个轴执行压辊动作@长有效 *)
    o_xManuConfirmSensorPos_LastAxis: BOOL; (* 最后一个轴手动确认传感器位置标志 *)

    (* 传感器电机运动 *)
    o_xSensorGoTargetPos_All: BOOL;      (* 所有轴向目标位置运动@到位后清除 *)
    o_rSenserTarPos_All: REAL;           (* 运动的目标位置 *)

    (* 动作控制 *)
    o_xExcuteAutoPreRegister_Ver: BOOL;  (* 执行纵向自动套印 *)
    o_xExcuteAutoPreRegisterDne_Ver: BOOL;(* 执行纵向自动套印完成 *)
    o_xExcuteAutoPreRegisterFailed_Ver: BOOL; (* 执行纵向自动套印失败 *)
    o_xAutoPreRegisterFinish_Ver: BOOL;  (* 执行纵向自动套印完成 *)
    o_byArcAdjAutoCtl: BYTE;             (* 套色手自动控制 *)

    (* 状态信息 *)
    o_eSts: EnumAutoPrintMasterStep;     (* 主状态机状态 *)
    o_iMsgInf: EnumAutoMaticRegisterCtlMsg; (* 信息 *)

    (* 轴控制输出 *)
    o_axAxisFindModuleEn: ARRAY[1..MAX_UNIT_NUM] OF BOOL; (* 轴寻找模块使能 *)
    o_axAxisCmd: ARRAY[1..MAX_UNIT_NUM] OF EnumFindCommand; (* 轴命令 *)

    (* 寻找结果 *)
 //   o_astFindResult: ARRAY[1..MAX_UNIT_NUM] OF StFindResult; (* 各轴寻找结果 *)
    o_xAllFindComplete: BOOL;            (* 所有轴寻找完成 *)

    (* 调整量输出 *)
    o_arAdjValue_Point: ARRAY[1..MAX_UNIT_NUM] OF REAL; (* 调整量@点 *)
    o_axAxisStartPress: ARRAY[1..MAX_UNIT_NUM] OF BOOL; (* 合压输出 *)
	o_arAdjPos_um	:ARRAY [1..MAX_UNIT_NUM] OF LREAL;(*色组调整了*)

    (* 流水线状态 *)
    o_iCurrentAxisIndex: INT;            (* 当前处理的轴索引（从后往前） *)
    o_xCurrentAxisProcessing: BOOL;      (* 当前轴正在处理 *)

    (* 轴状态显示 *)
    o_eState: ARRAY[1..MAX_UNIT_NUM] OF EnumFindState; (* 各轴状态描述 *)
	o_iErrorCode: ARRAY[1..MAX_UNIT_NUM] OF EnumFindState; (* 各轴报错*)
END_VAR
VAR
    (* 主状态机 *)
    eMainSts: EnumAutoPrintMasterStep;
    iMsgInf: EnumAutoMaticRegisterCtlMsg;

    (* 准备阶段变量 *)
    fbTimeOutTon: TON;                   (* 超时计时器 *)
    iLastAxisId: INT;                    (* 最后一个轴id *)
    rWaitFilmLenth: REAL;                (* 等待的料长@m *)
    xCheckSensorToTargetPos: BOOL;       (* 检查传感器到达目标位置 *)
    rTmp: REAL;                          (* 临时变量 *)
    xTmp: BOOL;                          (* 临时布尔 *)

    (* 传感器相关 *)
    axRollerPressSts_In: ARRAY[1..MAX_UNIT_NUM] OF BOOL; (* 压辊状态 *)
    axSensorMotorIdle: ARRAY[1..MAX_UNIT_NUM] OF BOOL;   (* 传感器电机空闲 *)

    (* 寻找结果 *)
 //   astFindResult: ARRAY[1..MAX_UNIT_NUM] OF StFindResult;

    (* 控制标志 *)
    xNextStep: BOOL;                     (* 初始化完成 *)

    (* 轴间关系 *)
    aiBeforeAxisId: ARRAY[1..MAX_UNIT_NUM] OF INT; (* 前轴号 *)
    aiAfterAxisId: ARRAY[1..MAX_UNIT_NUM] OF INT;  (* 后轴号 *)

    (* 临时变量 *)
    iN: INT;
	iM:INT;
    iAxisId: INT;
	iAxisId_Calc :INT;
    iBeforeAxisId: INT;
    iAfterAxisId: INT;

    pstStGrpParam_Save: POINTER TO StGrpParam_Save;
    pstStUnitParam_Save: POINTER TO StUnitParam_Save;
    pstStRSV_UnitParam_UnSave: POINTER TO StRSV_UnitParam_UnSave;
    pstStRSV_GrpParam_Save: POINTER TO StRSV_GrpParam_Save;

    rGirth: REAL;
    rFilmLength: REAL;

    (* 寻找结果存储 *)
    aiCurBestSignalPos: ARRAY[1..MAX_UNIT_NUM] OF INT;  (* 当前色最佳位置 *)
    aiPreLabelPos: ARRAY[1..MAX_UNIT_NUM] OF INT;       (* 前色位置 *)

    (* 轴命令控制 *)
    axAxisCmdSingle: ARRAY[1..MAX_UNIT_NUM] OF BOOL;    (* 轴单色命令触发 *)
    axAxisCmdMix: ARRAY[1..MAX_UNIT_NUM] OF BOOL;       (* 轴混色命令触发 *)

    (* 新增：简化流水线状态管理 *)
    axAxisComplete: ARRAY[1..MAX_UNIT_NUM] OF BOOL;     (* 轴完成标志 *)
    axAxisNeedPress: ARRAY[1..MAX_UNIT_NUM] OF BOOL;    (* 轴需要合压标志 *)
    axAxisPressDone: ARRAY[1..MAX_UNIT_NUM] OF BOOL;    (* 轴合压完成标志 *)
    axAxisStartPressTriggered: ARRAY[1..MAX_UNIT_NUM] OF BOOL; (* 轴合压已触发标志 *)

    (* 新增：前轴合压请求记录 *)
    axBeforeAxisPressRequested: ARRAY[1..MAX_UNIT_NUM] OF BOOL; (* 前轴合压已请求 *)

    (* 新增：所有轴完成标志 *)
    xAllAxisComplete: BOOL;               (* 所有轴完成标志 *)
	xCalculationCompleted:BOOL;           (*所有轴调整量计算完成*)

    (* 新增：轴状态描述数组 *)
  //  asAxisStatus: ARRAY[1..MAX_UNIT_NUM] OF STRING(50); (* 各轴状态描述 *)

    (* 新增：第一轴合压完成标志 *)
    xFirstAxisPressComplete: BOOL;        (* 第一轴合压完成 *)

	(*快速调整计算*)
	iIndexTmp:INT;(*//临时索引*)
	iIndex1TO2:INT;(*//从前向后的当前索引*)
	iIndex2TO1:INT;(*//从后向前的当前索引*)
	iAxisNum_1TO2:INT;(*//从前向后轴个数*)
	aiAxisIdList_FastAdj_1TO2:ARRAY [1..MAX_UNIT_NUM] OF INT;(*//从前到后压辊轴id*)
	iAxisNum_2TO1:INT;(*//从后向前轴个数*)
	aiAxisIdList_FastAdj_2TO1:ARRAY [1..MAX_UNIT_NUM] OF INT;(*//从后向前压辊轴id*)
	xCanFastAdj:BOOL;(*//可以快速对版标志*)
	iNeedFastAdjAxisNum:INT;(*//需要快速对版轴个数*)
	axFastAdjing:ARRAY [1..MAX_UNIT_NUM] OF BOOL;(*//快速对版中*)
	iAxisIdTmp:INT;
	axAdjust_ing: ARRAY [1..MAX_UNIT_NUM] OF BOOL;
	axAdjust_finish: ARRAY [1..MAX_UNIT_NUM] OF BOOL;
	xAllAdjust_finish:BOOL;
	byMeanANDAutoChangeCnt:BYTE;

END_VAR

{IMPLEMENTATION}
(* 初始化输出 *)
o_xAlarm := FALSE;
//o_xWaitingFilmLenthEn := FALSE;
o_xAutoPreRegister_Hor := FALSE;
o_xManuConfirmSensorPos_LastAxis := FALSE;
o_xSensorGoTargetPos_All := FALSE;
o_rSenserTarPos_All := 0;
o_xExcuteAutoPreRegister_Ver := FALSE;
o_xExcuteAutoPreRegisterDne_Ver := FALSE;
o_xExcuteAutoPreRegisterFailed_Ver := FALSE;
o_xAutoPreRegisterFinish_Ver := FALSE;
o_byArcAdjAutoCtl := 0;
o_xAllFindComplete := FALSE;
o_eSts := APM_STEP_IDLE;
o_iMsgInf := AMRC_MSG_NORMAL;
o_iCurrentAxisIndex := 0;
o_xCurrentAxisProcessing := FALSE;

FOR iN := 1 TO MAX_UNIT_NUM BY 1 DO
    o_axAxisFindModuleEn[iN] := FALSE;
    o_axAxisCmd[iN] := FIND_CMD_IDLE;
    i_pastFindResults^[iN].xSuccess := FALSE;
    i_pastFindResults^[iN].iErrorCode := 0;
   //
   // o_axAxisStartPress[iN] := FALSE;
  //  o_axAxisStatus[iN] := '';
END_FOR

(* 检查指针有效性 *)
IF i_pstStSysParam = 0 OR
   i_pastStIOMap_AxisBasic = 0 OR
   i_pastStAxisRapidAdjProf_V = 0 OR
   i_pafbKS_FB_AxisFindModule = 0 THEN
    RETURN;
END_IF

(* 获取外部状态 *)
FOR iN := 1 TO MAX_UNIT_NUM BY 1 DO
    pstStRSV_UnitParam_UnSave := ADR(i_pstStSysParam^.astStRSV_UnitParam_UnSave[iN]);
    axRollerPressSts_In[iN] := i_pastStIOMap_AxisBasic^[iN].o_xRel_Press;
    axSensorMotorIdle[iN] := pstStRSV_UnitParam_UnSave^.wState_FiberMove.8;
END_FOR

IF i_xEn THEN
    (* 前期准备阶段 *)
    rWaitFilmLenth := i_rMachineryFilmLenth ;  (* 等待机组料长等待 *)

    IF NOT o_xEning THEN
        (* 做参数初始化 *)
        o_xAlarm := FALSE;
        o_xAutoPreRegister_Hor := FALSE;
        o_xSensorGoTargetPos_All := FALSE;
        o_xManuConfirmSensorPos_LastAxis := FALSE;
        o_rSenserTarPos_All := 0;
        o_xExcuteAutoPreRegister_Ver := FALSE;
        o_xAutoPreRegisterFinish_Ver := FALSE;
       // o_xWaitingFilmLenthEn := FALSE;
        o_byArcAdjAutoCtl := 2;  (* 套色手动 *)

        fbTimeOutTon(IN:=FALSE);
        iLastAxisId := 0;
        xCheckSensorToTargetPos := FALSE;

        (* 计算最后一个轴ID *)
        IF i_byAxisNum > 0 AND i_byAxisNum <= MAX_UNIT_NUM THEN
            iLastAxisId := i_aiAxisList[i_byAxisNum];
        END_IF

        (* 初始化寻找结果 *)
        FOR iN := 1 TO MAX_UNIT_NUM BY 1 DO
            i_pastFindResults^[iN].xSuccess := FALSE;
            i_pastFindResults^[iN].iErrorCode := 0;
			o_arAdjValue_Point[iN] := 0.0;
			o_arAdjPos_um[iN] := 0.0;
			(* 初始化状态标志 *)
            axAxisComplete[iN] := FALSE;
            axAxisNeedPress[iN] := FALSE;
            axAxisPressDone[iN] := FALSE;
            axAxisStartPressTriggered[iN] := FALSE;
            axBeforeAxisPressRequested[iN] := FALSE;
            axAxisCmdSingle[iN] := FALSE;
            axAxisCmdMix[iN] := FALSE;
			//2026.05.19.200017+
			axAdjust_ing[iN]:=FALSE;
			axFastAdjing[iN]:=FALSE;
			axAdjust_finish[iN]:=FALSE;
        END_FOR

        (* 初始化轴间关系 *)
        FOR iN := 1 TO i_byAxisNum BY 1 DO
            iAxisId := i_aiAxisList[iN];

            (* 计算前后轴关系 *)
            IF iN = 1 THEN
                (* 第一个轴 *)
                aiBeforeAxisId[iAxisId] := -1;
                aiAfterAxisId[iAxisId] := i_aiAxisList[2];
            ELSIF iN = i_byAxisNum THEN
                (* 最后一个轴 *)
                aiBeforeAxisId[iAxisId] := i_aiAxisList[i_byAxisNum-1];
                aiAfterAxisId[iAxisId] := -1;
            ELSE
                (* 中间轴 *)
                aiBeforeAxisId[iAxisId] := i_aiAxisList[iN-1];
                aiAfterAxisId[iAxisId] := i_aiAxisList[iN+1];
            END_IF
		   //o_axAxisStartPress[iAxisId] := TRUE;
          //  asAxisStatus[iAxisId] := '空闲';
        END_FOR
		xNextStep:=TRUE;
		FOR iN:=2 TO i_byAxisNum BY 1 DO(*开始的时候全部打手动*)
			iAxisId:= i_aiAxisList[iN];
			pstStUnitParam_Save:= ADR(i_pstStsysParam^.astStUnitParam_Save[iAxisId]);
			IF pstStUnitParam_Save^.dwFlag_Sts.0 OR pstStUnitParam_Save^.dwFlag_Sts.1 THEN
				pstStUnitParam_Save^.dwFlag_Sts.0:= FALSE;
				pstStUnitParam_Save^.dwFlag_Sts.1:= FALSE;
				xNextStep:=FALSE;
			END_IF
		END_FOR
        (* 初始化全自动控制变量 *)
        xAllAxisComplete := FALSE;
        xFirstAxisPressComplete := FALSE;
		xCanFastAdj:=FALSE;

        IF xNextStep THEN
			o_xEning := TRUE;
			eMainSts := APM_STEP_TIPS;
			iMsgInf := AMRC_MSG_NORMAL;
		END_IF
      //  xInitDone := FALSE;
    END_IF

    (* 主状态机处理 - 前期准备阶段 *)
    CASE eMainSts OF
        APM_STEP_IDLE:
            (* 空闲状态 *)
            ;

        APM_STEP_TIPS:
            IF i_xTipsConfirm THEN
                eMainSts := APM_STEP_TIPS_ALARM;
            END_IF

        APM_STEP_TIPS_ALARM:
            o_xAlarm := TRUE;
            fbTimeOutTon(IN:=TRUE, PT:=T#3S);

            IF fbTimeOutTon.Q THEN
                IF i_xUseAutoPreRegister_Hor THEN
                    eMainSts := APM_STEP_AUTO_HOR;
                ELSE
                    IF i_xUseAutoSensorPos THEN
                        eMainSts := APM_STEP_AUTOSENSORPOS;
                    ELSE
                        eMainSts := APM_STEP_AUTO_VER;
                    END_IF
                END_IF
            END_IF

            (* 复位计时器 *)
            IF eMainSts <> APM_STEP_TIPS_ALARM THEN
                o_xAlarm := FALSE;
                fbTimeOutTon(IN:=FALSE);
            END_IF

        (* 横向动作状态处理 *)
        APM_STEP_AUTO_HOR:
            IF i_xAutoPreRegisterIdle_Hor THEN
                o_xAutoPreRegister_Hor := TRUE;

                IF i_xAutoPreRegistering_Hor THEN
                    eMainSts := APM_STEP_AUTOING_HOR;
                ELSE
                    fbTimeOutTon(IN:=TRUE, PT:=T#1S);
                    IF fbTimeOutTon.Q THEN
                        eMainSts := APM_STEP_TIMEOUT;
                    END_IF
                END_IF
            ELSE
                eMainSts := APM_STEP_ERR;
            END_IF

            (* 错误信息处理 *)
            IF eMainSts = APM_STEP_ERR THEN
                iMsgInf := AMRC_MSG_ERR_BUSY_HOR;
            END_IF
            IF eMainSts = APM_STEP_TIMEOUT THEN
                iMsgInf := AMRC_MSG_TIMEOUT_HOR;
            END_IF

            (* 退出case复位计时器 *)
            IF eMainSts <> APM_STEP_AUTO_HOR THEN
                o_xAutoPreRegister_Hor := FALSE;
                fbTimeOutTon(IN:=FALSE);
            END_IF

        APM_STEP_AUTOING_HOR:
            IF NOT i_xAutoPreRegistering_Hor THEN
                IF i_xUseAutoSensorPos THEN
                    eMainSts := APM_STEP_AUTOSENSORPOS;
                ELSE
                    eMainSts := APM_STEP_AUTO_VER;
                END_IF
            END_IF

        (* 自动sensor位置控制 *)
        APM_STEP_AUTOSENSORPOS:
            IF i_xUseSensorPos_3rd THEN
                eMainSts := APM_STEP_SENSORPOSBYSYS3RD;
            ELSE
                eMainSts := APM_STEP_SENSORPOSBYMANU;
            END_IF

        (* 第三方设备获取传感器位置 *)
        APM_STEP_SENSORPOSBYSYS3RD:
            IF iLastAxisId <> 0 THEN
                IF NOT axRollerPressSts_In[iLastAxisId] THEN
					o_axAxisStartPress[iLastAxisId] := TRUE;
                    //o_xExcuteRollerPress_LastAxis := TRUE;
                END_IF
                eMainSts := APM_STEP_WAITPOSBY3RD;
            ELSE
                eMainSts := APM_STEP_ERR;
            END_IF

            IF eMainSts = APM_STEP_ERR THEN
                iMsgInf := AMRC_MSG_ERR_LASTAXISID_INVALID;
            END_IF

        APM_STEP_WAITPOSBY3RD:
            IF NOT i_xSensorPosValid_3rd THEN
                eMainSts := APM_STEP_SENSOR_TO_TARGETPOS;
                o_rSenserTarPos_All := i_rSenserPos_3rd;
            ELSE
                IF i_rVel <> 0 THEN
                    rTmp := rWaitFilmLenth / i_rVel * 60;
                ELSE
                    rTmp := rWaitFilmLenth / 30.0 * 60;
                END_IF
                rTmp := rTmp * 1000;  (* 转换为毫秒 *)

                fbTimeOutTon(IN:=TRUE, PT:=REAL_TO_TIME(rTmp));
                IF fbTimeOutTon.Q THEN
                    eMainSts := APM_STEP_TIMEOUT;
                END_IF
            END_IF

            (* 输出信息 *)
            IF eMainSts = APM_STEP_TIMEOUT THEN
                iMsgInf := AMRC_MSG_TIMEOUT_WAITPOS_3RD;
            END_IF

            IF eMainSts <> APM_STEP_WAITPOSBY3RD THEN
                fbTimeOutTon(IN:=FALSE);
            END_IF

        (* 手动确认传感器位置 *)
        APM_STEP_SENSORPOSBYMANU:
            IF iLastAxisId <> 0 THEN
                IF NOT axRollerPressSts_In[iLastAxisId] THEN
					o_axAxisStartPress[iLastAxisId] := TRUE;
                    //o_xExcuteRollerPress_LastAxis := TRUE;
                END_IF
                eMainSts := APM_STEP_WAITPOSBYMANU;
            ELSE
                eMainSts := APM_STEP_ERR;
            END_IF

            IF eMainSts = APM_STEP_ERR THEN
                iMsgInf := AMRC_MSG_ERR_LASTAXISID_INVALID;
            END_IF

        APM_STEP_WAITPOSBYMANU:
            o_xManuConfirmSensorPos_LastAxis := TRUE;

            IF  i_xSensorPosValid_Manu THEN
                eMainSts := APM_STEP_SENSOR_TO_TARGETPOS;
                o_rSenserTarPos_All := i_rSensorPos_Manu;
            ELSE
                IF i_rVel <> 0 THEN
                    rTmp := rWaitFilmLenth / i_rVel * 60;
                ELSE
                    rTmp := rWaitFilmLenth / 30.0 * 60;;
                END_IF
                rTmp := rTmp * 1000;  (* 转换为毫秒 *)

                fbTimeOutTon(IN:=TRUE, PT:=REAL_TO_TIME(rTmp));
                IF fbTimeOutTon.Q THEN
                    eMainSts := APM_STEP_TIMEOUT;
                END_IF
            END_IF

            (* 输出信息 *)
            IF eMainSts = APM_STEP_TIMEOUT THEN
                iMsgInf := AMRC_MSG_TIMEOUT_WAITPOS_MANU;
            END_IF

            IF eMainSts <> APM_STEP_WAITPOSBYMANU THEN
                fbTimeOutTon(IN:=FALSE);
                o_xManuConfirmSensorPos_LastAxis := FALSE;
            END_IF

        (* 传感器电机向目标位置运动 *)
        APM_STEP_SENSOR_TO_TARGETPOS:
            xTmp := KS_CheckSensorMotorIdleSts(0, i_byAxisNum, i_aiAxisList, axSensorMotorIdle);
            IF xTmp THEN
                o_xSensorGoTargetPos_All := TRUE;
            END_IF

            IF o_xSensorGoTargetPos_All THEN
				eMainSts := APM_STEP_SENSOR_TO_TARGETPOSING;
				o_xSensorGoTargetPos_All := FALSE;
            END_IF

        APM_STEP_SENSOR_TO_TARGETPOSING:
            xTmp := KS_CheckSensorMotorIdleSts(iLastAxisId, i_byAxisNum, i_aiAxisList, axSensorMotorIdle);

            IF i_xUseFindBestPosStep THEN
                xCheckSensorToTargetPos := TRUE;
                eMainSts := APM_STEP_AUTO_VER;
            ELSE
                IF xTmp THEN
                    eMainSts := APM_STEP_AUTO_VER;
                END_IF
            END_IF

        (* 纵向全自动套印 - 流水线处理 *)
        APM_STEP_AUTO_VER:
            (* 启动寻找模块 *)
            o_xExcuteAutoPreRegister_Ver := TRUE;
            o_xCurrentAxisProcessing := TRUE;
            axAxisNeedPress[iLastAxisId]:=TRUE;
            eMainSts := APM_STEP_AUTOING_VER;

        APM_STEP_AUTOING_VER:
            (* 简化流水线处理逻辑 - 只负责触发前轴合压和激活寻找模块 *)
            o_xCurrentAxisProcessing := TRUE;
            o_iCurrentAxisIndex := 0;

            (* 首先，更新所有轴的状态描述 *)
            xAllAxisComplete := TRUE;  (* 假设所有轴都完成 *)

            FOR iN := i_byAxisNum TO 1 BY -1 DO
                iAxisId := i_aiAxisList[iN];
                iBeforeAxisId := aiBeforeAxisId[iAxisId];

                (* 跳过已完成的轴 *)
                IF axAxisComplete[iAxisId] THEN
                    CONTINUE;
                END_IF

                (* 标记有轴未完成 *)
                xAllAxisComplete := FALSE;

                (* 记录当前正在处理的轴索引 *)
                IF NOT axAxisComplete[iAxisId] THEN
                    o_iCurrentAxisIndex := iN;
                END_IF

                (* 第一轴特殊处理：只需要合压 *)
                IF iN = 1 THEN
                    (* 第一轴尚未合压完成 *)
                    IF NOT axAxisPressDone[iAxisId] THEN
                        (* 检查是否需要合压 *)
                        IF axAxisNeedPress[iAxisId] AND NOT axAxisPressDone[iAxisId] THEN
                            (* 触发合压 *)
                            IF NOT axAxisStartPressTriggered[iAxisId] THEN
                                o_axAxisStartPress[iAxisId] := TRUE;
                                axAxisStartPressTriggered[iAxisId] := TRUE;
                              //  asAxisStatus[iAxisId] := '合压中';
                            END_IF

                            (* 检查合压是否完成 *)
                            IF axRollerPressSts_In[iAxisId] THEN
                                (* 合压完成 *)
                                o_axAxisStartPress[iAxisId] := FALSE;
                                axAxisPressDone[iAxisId] := TRUE;
                                axAxisComplete[iAxisId] := TRUE;
                             //   asAxisStatus[iAxisId] := '完成';
                                xFirstAxisPressComplete := TRUE;
                            END_IF
                        END_IF
                    END_IF
                    CONTINUE;
                END_IF

                (* 非第一轴的处理逻辑 *)

                (* 1. 检查是否需要合压 *)
                IF axAxisNeedPress[iAxisId] AND NOT axAxisPressDone[iAxisId] THEN
                    (* 需要合压但未合压 *)
                    IF NOT axAxisStartPressTriggered[iAxisId] THEN
                        (* 触发合压 *)
                        IF iN = i_byAxisNum THEN
                            (* 最后一个轴 *)
							o_axAxisStartPress[iLastAxisId] := TRUE;
                        ELSE
                            (* 其他轴 *)
                            o_axAxisStartPress[iAxisId] := TRUE;
                        END_IF
                        axAxisStartPressTriggered[iAxisId] := TRUE;
                     //   asAxisStatus[iAxisId] := '等待合压';
                    END_IF

                    (* 检查合压是否完成 *)
                    IF axRollerPressSts_In[iAxisId] THEN
                        (* 合压完成 *)
//                         IF iN = i_byAxisNum THEN
// 							o_axAxisStartPress[iLastAxisId] := TRUE;
//                         END_IF
                        o_axAxisStartPress[iAxisId] := FALSE;
                        axAxisPressDone[iAxisId] := TRUE;

                        (* 激活寻找模块并发送单色寻找命令 *)
                        o_axAxisFindModuleEn[iAxisId] := TRUE;
                        IF NOT axAxisCmdSingle[iAxisId] THEN
                            o_axAxisCmd[iAxisId] := FIND_CMD_START_SINGLE;
                            axAxisCmdSingle[iAxisId] := TRUE;
                        END_IF

                      //  asAxisStatus[iAxisId] := '寻找单色中';
                    END_IF
                END_IF

                (* 2. 检查轴寻找模块的状态 *)
                IF axAxisPressDone[iAxisId] AND NOT axAxisComplete[iAxisId] THEN
                    (* 轴已合压完成，正在寻找中 *)

                    (* 激活寻找模块 *)
                    o_axAxisFindModuleEn[iAxisId] := TRUE;

                    (* 3. 检查是否需要触发前轴合压 *)
                    IF iBeforeAxisId <> -1 THEN
                        (* 检查轴寻找模块是否发出前轴合压信号 *)
                        IF i_pafbKS_FB_AxisFindModule^[iAxisId].o_xBeforeAxisStartPress AND
                           NOT axBeforeAxisPressRequested[iAxisId] THEN
                            (* 触发前轴合压 *)
                            axAxisNeedPress[iBeforeAxisId] := TRUE;
                            axBeforeAxisPressRequested[iAxisId] := TRUE;
                        END_IF
                    END_IF

                    (* 4. 检查轴是否完成 *)
                    IF i_pafbKS_FB_AxisFindModule^[iAxisId].o_xDone THEN
                        (* 轴寻找完成 *)
                        o_axAxisFindModuleEn[iAxisId] := FALSE;
                        axAxisComplete[iAxisId] := TRUE;

                        (* 保存寻找结果 *)
                        i_pastFindResults^[iAxisId] := i_pafbKS_FB_AxisFindModule^[iAxisId].o_stResult;
                        aiCurBestSignalPos[iAxisId] := i_pastFindResults^[iAxisId].iCurBestPos;

                        (* 记录前色位置（如果找到混色）*)
                        IF i_pastFindResults^[iAxisId].iPreLabelPos >= 0 THEN
                            aiPreLabelPos[iAxisId] := i_pastFindResults^[iAxisId].iPreLabelPos;
                        END_IF

                        (* 复位命令 *)
                        IF axAxisCmdSingle[iAxisId] THEN
                            o_axAxisCmd[iAxisId] := FIND_CMD_IDLE;
                            axAxisCmdSingle[iAxisId] := FALSE;
                        END_IF

                        IF axAxisCmdMix[iAxisId] THEN
                            o_axAxisCmd[iAxisId] := FIND_CMD_IDLE;
                            axAxisCmdMix[iAxisId] := FALSE;
                        END_IF
                    END_IF
                END_IF
            END_FOR

            (* 检查是否所有轴都完成 *)
            IF xAllAxisComplete THEN
                eMainSts := APM_STEP_CALC_ADJUSTMENTS;
                (* 复位全自动套印标志 *)
                o_xExcuteAutoPreRegister_Ver := FALSE;
                o_xAutoPreRegisterFinish_Ver := TRUE;
            END_IF

        APM_STEP_CALC_ADJUSTMENTS:
            (* 计算调整量 *)
           // o_xBusy := TRUE;

            (* 计算每个轴的调整量（从第二个轴开始）*)
            FOR iN := 2 TO i_byAxisNum BY 1 DO
                iAxisId := i_aiAxisList[iN];

                (* 获取参数指针 *)
                pstStUnitParam_Save := ADR(i_pstStSysParam^.astStUnitParam_Save[iAxisId]);
                pstStGrpParam_Save := ADR(i_pstStSysParam^.astStGrpParam_Save);

                (* 计算纵向调整量 *)
                IF aiCurBestSignalPos[iAxisId] >= 0 AND aiPreLabelPos[iAxisId] >= 0 THEN
                    o_arAdjValue_Point[iAxisId] := KS_CalculateVerticalAdjustment(
                        iAxisId,
                        aiCurBestSignalPos[iAxisId],
                        aiPreLabelPos[iAxisId],
                        pstStUnitParam_Save,
                        pstStGrpParam_Save
                    );
                ELSE
                    o_arAdjValue_Point[iAxisId] := 0.0;
                END_IF
            END_FOR
            xCalculationCompleted:=FALSE;
			(*动作执行*)

			FOR iN:=2 TO i_byAxisNum BY 1 DO
				iAxisId:=i_aiAxisList[iN];
				pstStUnitParam_Save:= ADR(i_pstStsysParam^.astStUnitParam_Save[iAxisId]);
				o_arAdjPos_um[iAxisId]:=0;
				FOR iM:=2 TO iN BY 1 DO
					iAxisId_Calc:= i_aiAxisList[iM];
					(*当前色获取到的粗采样点数*)
					rTmp:=o_arAdjValue_Point[iAxisId_Calc];(*记录位置*)
					(*累加@此时单位还是粗采样点数*)
					o_arAdjPos_um[iAxisId]:=o_arAdjPos_um[iAxisId] + rTmp;
				END_FOR
				(*测试*)
				//o_arAdjPos_um[iAxisId]:=15000*iAxisId;
				(*2026.3.26.213041+ by liu.yt*)
				(*将调整的粗采样点数转换到+-MAX_ROUNDSAMPLE_NUM/2范围内*)
				WHILE o_arAdjPos_um[iAxisId] < -MAX_ROUNDSAMPLE_NUM / 2 DO
					o_arAdjPos_um[iAxisId] := o_arAdjPos_um[iAxisId] + MAX_ROUNDSAMPLE_NUM;
				END_WHILE
				WHILE o_arAdjPos_um[iAxisId] > MAX_ROUNDSAMPLE_NUM / 2 DO
					o_arAdjPos_um[iAxisId] := o_arAdjPos_um[iAxisId] - MAX_ROUNDSAMPLE_NUM;
				END_WHILE(*此时单位还是粗采样点数*)
				(*计算um单位*)
				o_arAdjPos_um[iAxisId]:= o_arAdjPos_um[iAxisId]* pstStUnitParam_Save^.rGirth_PrnRoller*1000 / MAX_ROUNDSAMPLE_NUM;
			END_FOR
			xCalculationCompleted:=TRUE;
            (* 进入快速调整步骤 *)
            eMainSts := APM_STEP_FAST_ADJUSTMENT;

        APM_STEP_FAST_ADJUSTMENT:
            (* 快速对版调整 *)
            //o_xBusy := TRUE;
			Action_Excute();
			IF xAllAdjust_finish THEN
				eMainSts := APM_STEP_COMPLETE;
				byMeanANDAutoChangeCnt:=0;
			END_IF
        APM_STEP_COMPLETE:
            (* 完成 *)
           // o_xBusy := FALSE;
		   IF xAllAdjust_finish THEN(*全部调整完成-自动合压*)
			   xNextStep:=TRUE;
				FOR iN:=2 TO i_byAxisNum BY 1 DO(*开始的时候全部打手动*)
					iAxisId:= i_aiAxisList[iN];
					pstStUnitParam_Save:= ADR(i_pstStsysParam^.astStUnitParam_Save[iAxisId]);
					(*结束后全部打自动*)
					IF NOT pstStUnitParam_Save^.dwFlag_Sts.0 THEN
						pstStUnitParam_Save^.dwFlag_Sts.0:= TRUE;
						xNextStep:=FALSE;
					END_IF
				END_FOR
				IF xNextStep THEN
					o_xAllFindComplete := TRUE;
				END_IF

// 				byMeanANDAutoChangeCnt := byMeanANDAutoChangeCnt+1;
// 				IF  byMeanANDAutoChangeCnt < 3 THEN
// 					o_byArcAdjAutoCtl:=1;
// 					o_xWaitingFilmLenthEn := TRUE;
// 				ELSE
// 					o_xWaitingFilmLenthEn := FALSE;
//
// 					//xAllAdjust_finish:=FALSE;
// 				END_IF
			END_IF

        (* 超时步 *)
        APM_STEP_TIMEOUT:
            eMainSts := APM_STEP_ERR;
            iMsgInf := AMRC_MSG_TIMEOUT_HOR;

        (* 返回失败 *)
        APM_STEP_ERR:
            o_xExcuteAutoPreRegisterFailed_Ver := TRUE;
            o_xAllFindComplete := FALSE;
    END_CASE

    (* 调用所有轴的寻找模块 *)
    FOR iN := 1 TO i_byAxisNum BY 1 DO
        iAxisId := i_aiAxisList[iN];

        (* 获取参数指针 *)
        pstStRSV_UnitParam_UnSave := ADR(i_pstStSysParam^.astStRSV_UnitParam_UnSave[iAxisId]);
        pstStUnitParam_Save := ADR(i_pstStSysParam^.astStUnitParam_Save[iAxisId]);
        pstStGrpParam_Save := ADR(i_pstStSysParam^.astStGrpParam_Save);
        pstStRSV_GrpParam_Save := ADR(i_pstStSysParam^.astStRSV_GrpParam_Save);

        rGirth := pstStUnitParam_Save^.rGirth_PrnRoller;
        rFilmLength := pstStUnitParam_Save^.rFilmLengthFromPrevPressUnit;

        (* 获取前后轴号 *)
        iBeforeAxisId := aiBeforeAxisId[iAxisId];
        iAfterAxisId := aiAfterAxisId[iAxisId];

        (* 调用轴寻找模块 *)
        i_pafbKS_FB_AxisFindModule^[iAxisId](
            (* 基本输入 *)
            i_xEn := o_axAxisFindModuleEn[iAxisId],
            i_iAxisId := iAxisId,
            i_eCmd := o_axAxisCmd[iAxisId],
            i_xUseFindBestPosStep := i_xUseFindBestPosStep,

            (* 参数输入 *)
            i_pstStRSV_UnitParam_UnSave := pstStRSV_UnitParam_UnSave,
            i_pstStUnitParam_Save := pstStUnitParam_Save,
            i_pstStGrpParam_Save := pstStGrpParam_Save,
            i_rVel := i_rVel,
            i_rGirth := rGirth,
            i_rFilmLength := rFilmLength,
            i_iBeforeAxisId := iBeforeAxisId,
            i_iAfterAxisId := iAfterAxisId,
            i_rFindBestPos_MoveDis := pstStRSV_GrpParam_Save^.arFiberMove,

            (* 外部状态输入 *)
            i_xCoarseDone := axSensorMotorIdle[iAxisId],
            i_xPressDone := axRollerPressSts_In[iAxisId],
            i_xAutoMode := (eMainSts = APM_STEP_AUTOING_VER),
            i_xFind_IDLE := pstStRSV_UnitParam_UnSave^.byFlag_CommFromSlave.4,

            (* 开关参数 *)
            i_xSwitch_EnFastPress := pstStRSV_GrpParam_Save^.xSwitch_EnFastPress,
            i_xSwitch_RFailure := FALSE,
            i_xSwitch_FFailure := FALSE,
            i_xSpecialMarkEn := FALSE
        );

    END_FOR

ELSE
    (* 复位处理 *)
    IF o_xEning THEN
        o_xEning := FALSE;
        eMainSts := APM_STEP_IDLE;
        o_xAlarm := FALSE;
        o_xAutoPreRegister_Hor := FALSE;
        o_xManuConfirmSensorPos_LastAxis := FALSE;
        o_xSensorGoTargetPos_All := FALSE;
        o_rSenserTarPos_All := 0;
        o_xExcuteAutoPreRegister_Ver := FALSE;
      //  o_xWaitingFilmLenthEn := FALSE;
        xCheckSensorToTargetPos := FALSE;
        o_byArcAdjAutoCtl := 0;  (* 套色手动 *)
		xCalculationCompleted:=FALSE;
        (* 复位所有轴的寻找模块 *)
		FOR iN:=1 TO MAX_UNIT_NUM BY 1 DO
			 o_axAxisStartPress[iAxisId]:=FALSE;
		END_FOR
        FOR iN := 1 TO i_byAxisNum BY 1 DO
            iAxisId := i_aiAxisList[iN];
            (* 获取参数指针 *)
            pstStRSV_UnitParam_UnSave := ADR(i_pstStSysParam^.astStRSV_UnitParam_UnSave[iAxisId]);
            pstStUnitParam_Save := ADR(i_pstStSysParam^.astStUnitParam_Save[iAxisId]);
            pstStGrpParam_Save := ADR(i_pstStSysParam^.astStGrpParam_Save);
            pstStRSV_GrpParam_Save := ADR(i_pstStSysParam^.astStRSV_GrpParam_Save);

            rGirth := pstStUnitParam_Save^.rGirth_PrnRoller;
            rFilmLength := pstStUnitParam_Save^.rFilmLengthFromPrevPressUnit;

            (* 获取前后轴号 *)
            iBeforeAxisId := aiBeforeAxisId[iAxisId];
            iAfterAxisId := aiAfterAxisId[iAxisId];

            (* 调用轴寻找模块复位 *)
            i_pafbKS_FB_AxisFindModule^[iAxisId](
                (* 基本输入 *)
                i_xEn := TRUE,
                i_iAxisId := iAxisId,
                i_eCmd := FIND_CMD_RESET,
                i_xUseFindBestPosStep := i_xUseFindBestPosStep,

                (* 参数输入 *)
                i_pstStRSV_UnitParam_UnSave := pstStRSV_UnitParam_UnSave,
                i_pstStUnitParam_Save := pstStUnitParam_Save,
                i_pstStGrpParam_Save := pstStGrpParam_Save,
                i_rVel := i_rVel,
                i_rGirth := rGirth,
                i_rFilmLength := rFilmLength,
                i_iBeforeAxisId := iBeforeAxisId,
                i_iAfterAxisId := iAfterAxisId,
				i_rFindBestPos_MoveDis := pstStRSV_GrpParam_Save^.arFiberMove,

                (* 外部状态输入 *)
                i_xCoarseDone := pstStRSV_UnitParam_UnSave^.wState_FiberMove.8,
                i_xPressDone := axRollerPressSts_In[iAxisId],
                i_xAutoMode := FALSE,
                i_xFind_IDLE := pstStRSV_UnitParam_UnSave^.byFlag_CommFromSlave.4,

                (* 开关参数 *)
                i_xSwitch_EnFastPress := pstStRSV_GrpParam_Save^.xSwitch_EnFastPress,
                i_xSwitch_RFailure := i_xSwitch_RFailure,
                i_xSwitch_FFailure := i_xSwitch_FFailure,
                i_xSpecialMarkEn := FALSE
            );
			i_pastFindResults^[iAxisId] := i_pafbKS_FB_AxisFindModule^[iAxisId].o_stResult;
        END_FOR
    END_IF
END_IF

(* 输出状态 *)
o_eSts := eMainSts;
o_iMsgInf := iMsgInf;
//o_astFindResult := astFindResult;
g_axAutoFind_Press:=o_axAxisStartPress;
FOR iN := 1 TO i_byAxisNum BY 1 DO
	iAxisId := i_aiAxisList[iN];
	o_eState[iAxisId]:= i_pafbKS_FB_AxisFindModule^[iAxisId].o_eState;
	o_iErrorCode[iAxisId]:=i_pafbKS_FB_AxisFindModule^[iAxisId].o_stResult.iErrorCode;
END_FOR

//o_axAxisStatus := asAxisStatus;

(* ---- KS_FB_AxisFindModule.st ---- *)
(*@CES
Name=KS_FB_AxisFindModule
Type=FunctionBlock
TypeGuid=6f9dac99-8de1-4efc-8465-68ac443b7d08
Guid=fe608f45-03e0-4e2e-a249-20c440ac82a6
HasDeclaration=True
HasImplementation=True
*)
{DECLARATION}
FUNCTION_BLOCK KS_FB_AxisFindModule
VAR_INPUT
    (** 基本输入 **)
    i_xEn: BOOL;                         (** 模块使能 **)
    i_iAxisId: INT;                      (** 轴号 **)
    i_eCmd: EnumFindCommand;             (** 命令 **)
    i_xUseFindBestPosStep: BOOL;         (** 使用寻找最佳位置步骤 **)

    (** 参数输入 **)
    i_pstStRSV_UnitParam_UnSave: POINTER TO StRSV_UnitParam_UnSave; (** 单元参数 **)
    i_pstStUnitParam_Save: POINTER TO StUnitParam_Save; (** 单元参数 **)
    i_pstStGrpParam_Save: POINTER TO StGrpParam_Save; (** 组参数 **)
    i_rVel: REAL;                        (** 速度 **)
    i_rGirth: REAL;                      (** 版周长 **)
    i_rFilmLength: REAL;                 (** 料长 **)
    i_iBeforeAxisId: INT;                (** 前轴号 **)
    i_iAfterAxisId: INT;                 (** 后轴号 **)
    i_rFindBestPos_MoveDis: ARRAY [1..2] OF REAL; (** 光纤移动距离 **)

    (** 外部状态输入 **)
    i_xCoarseDone: BOOL;                 (** 粗调完成标志 **)
    i_xPressDone: BOOL;                  (** 合压完成标志 **)
    i_xAutoMode: BOOL;                   (** 自动模式标志 **)
    i_xFind_IDLE: BOOL;                  (** 当前轴全自动套印空闲 **)

    (** 开关参数 **)
    i_xSwitch_EnFastPress: BOOL;         (** 快速合压开关 **)
    i_xSwitch_RFailure: BOOL;            (** R失效开关 **)
    i_xSwitch_FFailure: BOOL;            (** F失效开关 **)
    i_xSpecialMarkEn: BOOL;              (** 特殊标使能 **)
END_VAR
VAR_OUTPUT
    (** 状态输出 **)
    o_eState: EnumFindState;             (** 当前状态 **)
    o_stResult: StFindResult;            (** 寻找结果 **)
    o_xBusy: BOOL;                       (** 忙标志 **)
    o_xDone: BOOL;                       (** 完成标志 **)
    o_xSuccess: BOOL;                    (** 成功标志 **)
    o_xError: BOOL;                      (** 错误标志 **)
    o_iErrorCode: INT;                   (** 错误代码 **)

    (** 控制输出 **)
    o_xNeedPress: BOOL;                  (** 需要合压 **)
    o_xBeforeAxisStartPress: BOOL;       (** 前轴开始合压（自动模式下使用）**)

    (** 从站控制信号 **)
    o_xFindFirstMark: BOOL;              (** 启动单色寻找@发送给从站 **)
    o_xFindPreMark: BOOL;                (** 启动混色寻找@发送给从站 **)
    o_xGateMoveFinish: BOOL;             (** 波门移动完成 **)
    o_xCurManuAdjust: BOOL;              (** 当前色需要手动调整 **)
    o_xPreCurManuAdjust: BOOL;           (** 前色需要手动调整 **)

    (** 光纤移动控制 **)
    o_xFiberMoveDisRunStart_FindSignal: BOOL; (** 光纤移动启动 **)
    o_rFiberMoveDistanceIn_FindSignal: REAL; (** 光纤移动距离 **)

    (** 参数设置输出 **)
    o_iGateSa: INT;                      (** 波门起始位置 **)

    (** 寻找状态标志 **)
    o_xSingleFound: BOOL;                (** 单色至少找到一次 **)
    o_xMixFound: BOOL;                   (** 混色找到 **)
    o_xHasAlarm: BOOL;                   (** 有报警 **)
	o_xHasAlarming: BOOL;                (** 有报警铃输出 **)
    o_xPressTriggered: BOOL;             (** 合压已触发（前轴）**)
END_VAR
VAR
    iN: INT;
    (** 状态机 **)
    eState: EnumFindState;
    ePrevState: EnumFindState;

    (** 寻找参数 **)
    byFindCycleCnt: BYTE;
    aiCurLabelPos: ARRAY[1..3] OF INT;
    arCurLabelWidth: ARRAY[1..3] OF REAL;
    rFiberMoveDist: ARRAY[1..2] OF REAL;
    iCurBestSignalPos: INT;

    (** 计时器 **)
    fbDelayTimer: TON;
    fbMixDelayTimer: TON;                (** 混色寻找延时计时器 **)
    iDelayTime: DINT;
    iTotalDelayTime: DINT;
    iMixDelayTime: DINT;                 (** 混色延时时间 **)

    (** 状态标志 **)
  //  xInitDone: BOOL;
    xCoarseChecked: BOOL;
    xGateAdjusted: BOOL;
	xMasterComplete:BOOL;				(*从站再找一次*)
	xMasterCompleteing:BOOL;			(*从站再找一次中*)
    xFindSingleSuccess: BOOL;            (** 单色寻找最终成功 **)
    xFindMixSuccess: BOOL;               (** 混色寻找最终成功 **)
    xFiberMoved: BOOL;
    xPressRequested: BOOL;
    xMixDelayStarted: BOOL;              (** 混色延时已开始 **)
    xFineAdjustStarted: BOOL;            (** 精调已开始 **)
    xFineAdjustComplete: BOOL;           (** 精调完成 **)

    (** 寻找结果标志 **)
    xSingleFoundAtLeastOnce: BOOL;       (** 单色至少找到一次 **)
    xMixFound: BOOL;                     (** 混色找到 **)
    xHasSingleError: BOOL;               (** 单色寻找有错误 **)
    xHasMixError: BOOL;                  (** 混色寻找有错误 **)

    (** 触发标志 **)
    xBeforeAxisPressTriggered: BOOL;     (** 前轴合压已触发标志 **)

    (** 错误处理 **)
    iErrorCount: INT;
	fbR_TRIG_HasAlarm :R_trig;
	fbTON_HasAlarming :TON;

    (** 临时变量 **)
    iTemp: INT;
    rTemp: REAL;

    pstStRSV_UnitParam_UnSave: POINTER TO StRSV_UnitParam_UnSave;
    pstStUnitParam_Save: POINTER TO StUnitParam_Save;
    pstStGrpParam_Save: POINTER TO StGrpParam_Save;

    (** 寻找延时 **)
    iFindSingleDelayTime: DINT;          (** 单色寻找延时@ms **)
    iFindMixDelayTime: DINT;             (** 混色寻找延时@ms **)

    (** 命令处理 **)
    eCmd: EnumFindCommand;
    xCmdRising: BOOL;
    xPrevCmd: EnumFindCommand;

    (** 寻找标志 **)
    xUseFindBestPosStep: BOOL;           (** 使用寻找最佳位置步骤 **)

    (** 从站计算精采样宽度 **)
    xFindMarkCenter_CalWidth: BOOL;
    xPreStsFineAdjFiber: BOOL;
    xStsFineAdjFiber: BOOL;

	iWaitFiberMoveDelayTime:DINT:=500;

	xNeedMsg:BOOL;
	sLogMsg: STRING;
	sTimeStamp_Tmp				: STRING;
	tChangeStsTime:TIME;
	tLastTime:TIME;
END_VAR
{IMPLEMENTATION}
IF i_pstStRSV_UnitParam_UnSave = 0 OR
   i_pstStUnitParam_Save = 0 OR
   i_pstStGrpParam_Save = 0 THEN
    RETURN;
END_IF

(** 初始化指针 **)
pstStRSV_UnitParam_UnSave := i_pstStRSV_UnitParam_UnSave;
pstStUnitParam_Save := i_pstStUnitParam_Save;
pstStGrpParam_Save := i_pstStGrpParam_Save;

(** 重置输出 **)
o_xBusy := FALSE;
o_xDone := FALSE;
o_xSuccess := FALSE;
o_xError := FALSE;
o_xNeedPress := FALSE;
o_xBeforeAxisStartPress := FALSE;
o_xGateMoveFinish := FALSE;
o_xCurManuAdjust := FALSE;
o_xPreCurManuAdjust := FALSE;
o_xFiberMoveDisRunStart_FindSignal := FALSE;
o_rFiberMoveDistanceIn_FindSignal := 0.0;
o_iGateSa := 0;
o_eState := eState;
o_xSingleFound := FALSE;
o_xMixFound := FALSE;
o_xHasAlarm := FALSE;
o_xPressTriggered := xBeforeAxisPressTriggered;

(** 保存设置 **)
xUseFindBestPosStep := i_xUseFindBestPosStep;

(** 检测沿信号 **)
xPrevCmd := eCmd;
eCmd := i_eCmd;
IF eCmd <> xPrevCmd THEN
    xCmdRising := TRUE;
ELSE
    xCmdRising := FALSE;
END_IF

IF i_xEn THEN

    (** 命令处理 **)
    IF xCmdRising THEN
        CASE eCmd OF
            FIND_CMD_START_SINGLE:
                IF eState = FIND_STATE_IDLE THEN
                    eState := FIND_STATE_INIT;
                 //   xInitDone := FALSE;
                    xFindSingleSuccess := FALSE;
                    xFindMixSuccess := FALSE;
                    o_stResult.xSuccess := FALSE;
                    xBeforeAxisPressTriggered := FALSE;  (** 重置触发标志 **)
                END_IF

            FIND_CMD_START_MIX:
                IF eState = FIND_STATE_IDLE OR eState = FIND_STATE_COMPLETE THEN
                    (** 直接进入混色寻找延时状态 **)
                    eState := FIND_STATE_DELAY_MIX;
                    xFindMixSuccess := FALSE;
                    o_stResult.xSuccess := FALSE;
                END_IF

            FIND_CMD_RESET:
                eState := FIND_STATE_IDLE;
              //  xInitDone := FALSE;
                xFindSingleSuccess := FALSE;
                xFindMixSuccess := FALSE;
                o_stResult.xSuccess := FALSE;
                o_xBusy := FALSE;
                o_xDone := TRUE;
                o_xSuccess := TRUE;
                o_xError := FALSE;
                o_xNeedPress := FALSE;
                o_xFindFirstMark := FALSE;
                o_xFindPreMark := FALSE;
                o_xGateMoveFinish := TRUE;
                o_xBeforeAxisStartPress := FALSE;
                xFindMarkCenter_CalWidth := FALSE;
                o_xFiberMoveDisRunStart_FindSignal := FALSE;
                xBeforeAxisPressTriggered := FALSE;
				xHasSingleError :=FALSE;
				xHasMixError:=FALSE;
				fbDelayTimer(iN:=FALSE);
				fbMixDelayTimer(iN:=FALSE);
				fbTON_HasAlarming(iN:=FALSE);
        END_CASE
    END_IF

	(*混色计时器挪到外面*)
	fbMixDelayTimer(IN:=xBeforeAxisPressTriggered, PT:=DINT_TO_TIME(iFindMixDelayTime));

    (** 状态机主循环 **)
    CASE eState OF
        FIND_STATE_IDLE:
            (** 空闲状态，等待命令 **)
            o_xBusy := FALSE;
            o_xDone := TRUE;
            o_xNeedPress := FALSE;

        FIND_STATE_INIT:
            (** 初始化寻找参数 **)
            o_xBusy := TRUE;
            (** 初始化参数 **)
            byFindCycleCnt := 0;
            FOR iTemp := 1 TO 3 BY 1 DO
                aiCurLabelPos[iTemp] := -1;
                arCurLabelWidth[iTemp] := 0.0;
            END_FOR

            FOR iN := 1 TO 3 BY 1 DO
                IF iN <= 2 THEN
                    g_aiCurLabelPos[i_iAxisId, iN] := -1;
                    g_arCurLabelWidth[i_iAxisId, iN] := 0.0;
                    g_rFiberMoveDist[i_iAxisId, iN] := 0;
                END_IF
                g_aiCurLabelPos[i_iAxisId, iN] := -1;
                g_arCurLabelWidth[i_iAxisId, iN] := 0.0;
            END_FOR
            iCurBestSignalPos := -1;
            xMixDelayStarted := FALSE;
            xFineAdjustStarted := FALSE;
            xFineAdjustComplete := FALSE;
            xFindMarkCenter_CalWidth := FALSE;
            xSingleFoundAtLeastOnce := FALSE;
            xMixFound := FALSE;
            xHasSingleError := FALSE;
            xHasMixError := FALSE;
            xBeforeAxisPressTriggered := FALSE;
			fbTON_HasAlarming(iN:=FALSE);
			fbR_TRIG_HasAlarm(clk:=FALSE);
			o_stResult.xSuccess := FALSE;
			o_stResult.iErrorCode := 0;

            (** 检查是否需要合压 **)
            IF i_iAfterAxisId = -1 AND i_xAutoMode THEN
                (** 最后一个轴，需要合压 **)
                o_xNeedPress := TRUE;
                eState := FIND_STATE_CHECK_COARSE;
            ELSE
                eState := FIND_STATE_CHECK_COARSE;
            END_IF

			(** 计算延时时间 **)
			IF i_rVel > 0 AND i_rGirth > 0 THEN
				(** 单色寻找前延时：等待1.5圈 **)
				iFindSingleDelayTime := REAL_TO_DINT(1.5 * 60.0 * i_rGirth / 1000.0 / i_rVel * 1000.0);

				(** 混色寻找延时 **)
				IF i_iBeforeAxisId <> -1 THEN
					iFindMixDelayTime := KS_CalculateMixFindDelayTime(
						i_iAxisId,
						i_iBeforeAxisId,
						pstStUnitParam_Save,
						i_rVel
					);
				END_IF
			ELSE
				iFindSingleDelayTime := 1000;  (** 默认1秒 **)
				iFindMixDelayTime := 30000;    (** 默认30秒 **)
			END_IF
			fbMixDelayTimer(IN:=FALSE);
        FIND_STATE_CHECK_COARSE:
            (** 检查粗调状态 **)
            o_xBusy := TRUE;
            IF i_xCoarseDone THEN
				IF i_iAfterAxisId = -1 AND i_xPressDone THEN
					(** 最后一个轴，且合压完成，不需要需要合压，直接进入找标 **)
					eState := FIND_STATE_DELAY_SINGLE;
				ELSE
					 xCoarseChecked := TRUE;
               		 eState := FIND_STATE_WAIT_PRESS;
				END_IF
            ELSE
                (** 粗调未完成，设置错误标志但不停止流程 **)
                xHasSingleError := TRUE;
                o_stResult.iErrorCode := FIND_ERR_COARSE_NOT_READY;
            END_IF

        FIND_STATE_WAIT_PRESS:
            (** 等待合压完成 **)
            o_xBusy := TRUE;

            IF i_xPressDone THEN
                o_xNeedPress := FALSE;
                xPressRequested := FALSE;
                (** 启动单色寻找前延时计时器 **)
                fbDelayTimer(IN:=TRUE, PT:=DINT_TO_TIME(iFindSingleDelayTime));
            ELSE
                o_xNeedPress := TRUE;
            END_IF

            IF fbDelayTimer.Q THEN
                fbDelayTimer(IN:=FALSE);
                eState := FIND_STATE_DELAY_SINGLE;
            END_IF

        FIND_STATE_DELAY_SINGLE:
            o_xBusy := TRUE;
            (** 等待从站空闲 **)
			IF i_xFind_IDLE THEN
				IF i_xAutoMode THEN(*自动模式*)
					(** 初始化从站参数 **)
					o_xFindFirstMark := TRUE;
					o_xCurManuAdjust := FALSE;
					eState := FIND_STATE_FIND_SINGLE;
				ELSE (*手动模式*)
					eState := FIND_STATE_FIND_SINGLE;
				END_IF
			END_IF
        FIND_STATE_FIND_SINGLE:
            (** 执行单色寻找 **)
            o_xBusy := TRUE;
            IF NOT i_xFind_IDLE THEN
				xMasterComplete:=FALSE;
			END_IF
			IF i_xAutoMode THEN(*自动模式*)
					(** 等待从站结果 从站状态机在7或者8时，表示该次寻找完成**)
				IF pstStRSV_UnitParam_UnSave^.byFlag_CommFromSlave.2 AND (pstStRSV_UnitParam_UnSave^.byMarkStep = 7
					OR pstStRSV_UnitParam_UnSave^.byMarkStep = 8)THEN
					(** 从站找标完成 **)
					o_xFindFirstMark := FALSE;

					(** 记录结果 **)
					IF pstStRSV_UnitParam_UnSave^.iCurLabelPos >= 0 THEN
						(** 找到标记 **)
						byFindCycleCnt := byFindCycleCnt + 1;
						aiCurLabelPos[byFindCycleCnt] := pstStRSV_UnitParam_UnSave^.iCurLabelPos;
						arCurLabelWidth[byFindCycleCnt] := pstStRSV_UnitParam_UnSave^.rGateSignalWidth_R;
						xSingleFoundAtLeastOnce := TRUE;  (** 标记至少找到一次 **)

						(** 快速合压模式：第一次找到就触发前轴合压 **)
						IF i_xAutoMode AND i_iBeforeAxisId <> -1 AND i_xSwitch_EnFastPress
						   AND byFindCycleCnt = 1 AND NOT xBeforeAxisPressTriggered THEN
							o_xBeforeAxisStartPress := TRUE;
							xBeforeAxisPressTriggered := TRUE;  (** 标记已触发 **)
						END_IF

						(** 如果使用最佳位置步骤且还没采完3次，继续采样 **)
						IF xUseFindBestPosStep AND byFindCycleCnt < 3 THEN
							eState := FIND_STATE_MOVE_FIBER;
						ELSE
							(** 采完3次或不使用最佳位置步骤 **)
							eState := FIND_STATE_CALC_BEST;
						END_IF
					ELSE
						(** 未找到标记，记录错误但不停止 **)
						//xHasSingleError := TRUE;
						o_stResult.iErrorCode := FIND_ERR_SINGLE_MARK_NOT_FOUND;
						o_xCurManuAdjust := TRUE;  (** 需要手动调整 **)

						(** 增加计数，继续尝试 **)
						byFindCycleCnt := byFindCycleCnt + 1;

						(** 如果还没采完3次，继续采样 **)
						IF xUseFindBestPosStep AND byFindCycleCnt < 3 THEN
							eState := FIND_STATE_MOVE_FIBER;
						ELSE
							(** 采完3次，进入下一步 **)
							eState := FIND_STATE_CALC_BEST;
						END_IF
					END_IF
				END_IF
			ELSE (*手动模式*)
				 (** 通过精采样计算当前波门内波形宽度 **)
				xFindMarkCenter_CalWidth := TRUE;
				xStsFineAdjFiber := pstStRSV_UnitParam_UnSave^.byFlag_CommFromSlave.3;
				(** 检查是否需要光纤精调 **)
				IF xUseFindBestPosStep AND NOT xPreStsFineAdjFiber AND xStsFineAdjFiber
				    AND pstStRSV_UnitParam_UnSave^.xFiberMoveIdle THEN
					xFindMarkCenter_CalWidth := FALSE;
					byFindCycleCnt := byFindCycleCnt + 1;
					(*手动模式，需要填写一个>=0的值作为波形的位置，保证后续逻辑正确，所以这里先填写一个波门位置，实际波形位置不在这里*)
					aiCurLabelPos[byFindCycleCnt] := pstStUnitParam_Save^.iGateSa;
					arCurLabelWidth[byFindCycleCnt] := pstStRSV_UnitParam_UnSave^.rWidth_FindMarkCenter;
					xSingleFoundAtLeastOnce := TRUE;  (** 标记至少找到一次 **)
					(** 如果使用最佳位置步骤且还没采完3次，继续采样 **)
					IF xUseFindBestPosStep AND byFindCycleCnt < 3 THEN
						eState := FIND_STATE_MOVE_FIBER;
					ELSE
						(** 采完3次或不使用最佳位置步骤 **)
						eState := FIND_STATE_CALC_BEST;
					END_IF
				END_IF
				xPreStsFineAdjFiber := xStsFineAdjFiber;
			END_IF
        FIND_STATE_MOVE_FIBER:
            (** 移动光纤到下一个采样位置 **)
            o_xBusy := TRUE;
             IF NOT i_xFind_IDLE THEN
				xMasterComplete:=FALSE;
			END_IF
            IF pstStRSV_UnitParam_UnSave^.xFiberMoveIdle THEN
                (** 计算移动距离 **)
                CASE byFindCycleCnt OF
                    1:  (** 第二次采样，左移3mm **)
                        rFiberMoveDist[1] := i_rFindBestPos_MoveDis[1];
                    2:  (** 第三次采样，右移6mm **)
                        rFiberMoveDist[1] := i_rFindBestPos_MoveDis[2];
                END_CASE

                (** 执行移动 **)
                o_rFiberMoveDistanceIn_FindSignal := rFiberMoveDist[1];
                o_xFiberMoveDisRunStart_FindSignal := TRUE;
                xMasterCompleteing:=FALSE;
                eState := FIND_STATE_WAIT_FIBER_MOVE;
            END_IF

        FIND_STATE_WAIT_FIBER_MOVE:
            (** 等待光纤移动完成 **)
            o_xBusy := TRUE;
             IF NOT i_xFind_IDLE THEN
				xMasterComplete:=FALSE;
			END_IF

            IF pstStRSV_UnitParam_UnSave^.xFiberMoveIdle THEN
               	o_xFiberMoveDisRunStart_FindSignal := FALSE;
				IF i_xAutoMode THEN(*自动模式*)
					(** 等待从站空闲 **)
					IF i_xFind_IDLE AND NOT xMasterCompleteing THEN
						xMasterCompleteing:=TRUE;
						xMasterComplete := TRUE;
					END_IF
					IF NOT i_xFind_IDLE AND xMasterCompleteing THEN
						 eState := FIND_STATE_FIND_SINGLE;
					END_IF
				ELSE (*手动模式*)
					 eState := FIND_STATE_FIND_SINGLE;
				END_IF
            END_IF
        FIND_STATE_CALC_BEST:
            (** 计算最佳位置 **)
            o_xBusy := TRUE;
            xMasterComplete := FALSE;
			(** 使用寻找最佳位置步骤，且至少找到过一次 **)
			KS_CalBestFiberMoveDisByRS(
				arCurLabelWidth,
				aiCurLabelPos,
				pstStGrpParam_Save^.byTriMark_SideB,
				pstStGrpParam_Save^.byTriMark_SideC,
				pstStGrpParam_Save^.iMarkTypeId,
				ADR(iCurBestSignalPos),
				ADR(rFiberMoveDist[1])
			);
            IF xSingleFoundAtLeastOnce AND xUseFindBestPosStep THEN
                IF iCurBestSignalPos <> -1 THEN
                    (** 计算成功 **)
					 xFindSingleSuccess := TRUE;
					o_stResult.iCurBestPos := iCurBestSignalPos;

					(** 移动光纤到最佳位置 **)
					IF pstStRSV_UnitParam_UnSave^.xFiberMoveIdle THEN
						o_rFiberMoveDistanceIn_FindSignal := rFiberMoveDist[1];
						o_xFiberMoveDisRunStart_FindSignal := TRUE;
						IF i_xSwitch_RFailure THEN
							o_xFiberMoveDisRunStart_FindSignal := FALSE;
						END_IF
						eState := FIND_STATE_ADJUST_GATE;
					END_IF
                ELSE
                    (** 计算失败，记录错误但继续流程 **)
                    xHasSingleError := TRUE;
                    o_stResult.iErrorCode := FIND_ERR_CALC_BEST_FAILED;
                    o_xCurManuAdjust := TRUE;  (** 需要手动调整 **)
                   // eState := FIND_STATE_ADJUST_GATE;  (** 继续流程 **)
                END_IF
            ELSE
                (** 没有找到单色或不使用最佳位置步骤 **)
                IF xSingleFoundAtLeastOnce THEN
                    (** 至少找到过一次，使用第一次采样的位置 **)
                    iCurBestSignalPos := aiCurLabelPos[1];
                    rFiberMoveDist[1] := rFiberMoveDist[1];  (** 移动回原原位 **)
					o_xFiberMoveDisRunStart_FindSignal := TRUE;
                    xFindSingleSuccess := TRUE;
                    o_stResult.iCurBestPos := iCurBestSignalPos;
                ELSE
                    (** 一次都没找到，不设置最佳位置 **)
					o_rFiberMoveDistanceIn_FindSignal := rFiberMoveDist[1];
                    o_xFiberMoveDisRunStart_FindSignal := TRUE;
                    iCurBestSignalPos := -1;
                    xHasSingleError := TRUE;
                END_IF
            END_IF
		 	(** 非快速合压模式：在当前轴处理完成后触发前轴合压 **)
			IF i_xAutoMode AND i_iBeforeAxisId <> -1 AND NOT xBeforeAxisPressTriggered THEN
				o_xBeforeAxisStartPress := TRUE;
				xBeforeAxisPressTriggered := TRUE;  (** 标记已触发 **)
				eState := FIND_STATE_ADJUST_GATE;  (** 继续流程 **)
			END_IF
        FIND_STATE_ADJUST_GATE:
            (** 调整波门位置 **)
            o_xBusy := TRUE;

            (** 等待光纤移动完成（如果有移动）**)
            IF pstStRSV_UnitParam_UnSave^.xFiberMoveIdle THEN
                o_xFiberMoveDisRunStart_FindSignal := FALSE;

                (** 如果单色找到 且为自动模式，设置波门位置；否则波门保持原位 **)
                IF xSingleFoundAtLeastOnce AND i_xAutoMode AND iCurBestSignalPos <> -1 THEN
                    (** 设置波门中心位置 **)
                    o_iGateSa := iCurBestSignalPos - pstStUnitParam_Save^.iGateWidthRoundPoints / 2;

                    (** 边界检查 **)
                    IF o_iGateSa < 0 THEN
                        o_iGateSa := o_iGateSa + 4000;
                    ELSIF o_iGateSa > 3999 THEN
                        o_iGateSa := o_iGateSa - 4000;
                    END_IF
					pstStUnitParam_Save^.iGateSa:= o_iGateSa;
                ELSE
                    (** 单色没找到或者手动模式，波门保持原位 **)
                   o_iGateSa:=pstStUnitParam_Save^.iGateSa;
                END_IF
                o_xGateMoveFinish := TRUE;

                IF xSingleFoundAtLeastOnce AND iCurBestSignalPos <> -1 THEN
                    o_stResult.iCurLabelPos := iCurBestSignalPos;
                ELSE
                    o_stResult.iCurLabelPos := -1;
                END_IF

                (** 检查是否需要寻找混色 因为手动模式设置前色轴位-1，所以直接完成，不需要处理**)
                IF i_iBeforeAxisId <> -1 THEN
                    (** 有前轴，需要寻找混色 **)
					IF  pstStUnitParam_Save^.iGateSa =o_iGateSa THEN
						eState := FIND_STATE_DELAY_MIX;
					END_IF
                ELSE
                    (** 没有前轴，完成 **)
                    eState := FIND_STATE_COMPLETE;
                END_IF
            END_IF

        FIND_STATE_DELAY_MIX:
            (** 混色寻找前延时 **)
            o_xBusy := TRUE;

            (** 启动混色延时计时器 **)
            IF NOT xMixDelayStarted THEN
                xMixDelayStarted := TRUE;
				//fbMixDelayTimer(IN:=FALSE);
            END_IF
          //  fbMixDelayTimer(IN:=xMixDelayStarted, PT:=DINT_TO_TIME(iFindMixDelayTime));
            (** 光纤精调 **)
			IF  NOT xFineAdjustStarted THEN
				 xFindMarkCenter_CalWidth := TRUE;
			END_IF
            xStsFineAdjFiber := pstStRSV_UnitParam_UnSave^.byFlag_CommFromSlave.3;

            (** 检查是否需要光纤精调 **)
            IF xUseFindBestPosStep AND NOT xPreStsFineAdjFiber AND xStsFineAdjFiber AND
               NOT xFineAdjustStarted AND pstStRSV_UnitParam_UnSave^.xFiberMoveIdle AND
               NOT fbMixDelayTimer.Q THEN
			    xFindMarkCenter_CalWidth := FALSE;
                eState := FIND_STATE_FINE_ADJUST;
            END_IF

            xPreStsFineAdjFiber := xStsFineAdjFiber;

            (** 检查混色延时是否结束 **)
            IF fbMixDelayTimer.Q THEN
                fbMixDelayTimer(IN:=FALSE);
                xMixDelayStarted := FALSE;
                o_xFindPreMark := TRUE;
                eState := FIND_STATE_FIND_MIX;
            END_IF

        FIND_STATE_FINE_ADJUST:
            (** 光纤精调 **)
            o_xBusy := TRUE;

            IF NOT xFineAdjustStarted THEN
                (** 计算精调距离 **)
                KS_CalBestFiberMoveDisByPS(
                    ADR(pstStRSV_UnitParam_UnSave^.rWidth_FindMarkCenter),
                    pstStGrpParam_Save^.byTriMark_SideB,
                    pstStGrpParam_Save^.byTriMark_SideC,
                    pstStGrpParam_Save^.iMarkTypeId,
                    ADR(rFiberMoveDist[2])
                );

                (** 执行精调移动 **)
                o_rFiberMoveDistanceIn_FindSignal := rFiberMoveDist[2];
                o_xFiberMoveDisRunStart_FindSignal := TRUE;
				IF i_xSwitch_FFailure THEN
					 o_xFiberMoveDisRunStart_FindSignal := FALSE;
				END_IF
                xFineAdjustStarted := TRUE;
                eState := FIND_STATE_WAIT_FINE_ADJ;
            END_IF

        FIND_STATE_WAIT_FINE_ADJ:
            (** 等待精调完成 **)
            o_xBusy := TRUE;
         //   fbMixDelayTimer(IN:=xMixDelayStarted, PT:=DINT_TO_TIME(iFindMixDelayTime));
            IF pstStRSV_UnitParam_UnSave^.xFiberMoveIdle THEN
                o_xFiberMoveDisRunStart_FindSignal := FALSE;
                xFineAdjustComplete := TRUE;

                (** 返回等待混色状态，继续等待混色延时 **)
                eState := FIND_STATE_DELAY_MIX;
            END_IF
			 (** 检查混色延时是否结束 **)
            IF fbMixDelayTimer.Q THEN
                fbMixDelayTimer(IN:=FALSE);
                xMixDelayStarted := FALSE;
                o_xFindPreMark := TRUE;
                eState := FIND_STATE_FIND_MIX;
            END_IF

        FIND_STATE_FIND_MIX:
            (** 执行混色寻找 **)
            o_xBusy := TRUE;

            (** 等待从站结果 **)
            IF pstStRSV_UnitParam_UnSave^.xFlag_FindPreSuccess THEN
                (** 记录前色位置 **)
                IF pstStRSV_UnitParam_UnSave^.iPreLabelPos >= 0 AND pstStRSV_UnitParam_UnSave^.iPreLabelPos < 4000 THEN
                    xMixFound := TRUE;
                    xFindMixSuccess := TRUE;
                    o_stResult.iPreLabelPos := pstStRSV_UnitParam_UnSave^.iPreLabelPos;
                ELSE
                    (** 前色位置无效 **)
                    xHasMixError := TRUE;
                    o_stResult.iErrorCode := FIND_ERR_PRE_POS_INVALID;
                    o_xPreCurManuAdjust := TRUE;  (** 需要手动调整 **)
                END_IF

                o_xFindPreMark := FALSE;
                eState := FIND_STATE_COMPLETE;
            END_IF

        FIND_STATE_COMPLETE:
            (** 寻找完成 **)
            o_xBusy := FALSE;
            o_xDone := TRUE;

            (** 设置最终成功标志：单色和混色都找到才算成功 **)
            IF i_iBeforeAxisId = -1 THEN
                (** 第一色，不需要寻找，只要合压完成就算成功 **)
                o_xSuccess := TRUE;
            ELSE
                (** 非第一色，需要单色和混色都找到 **)
                o_xSuccess := xSingleFoundAtLeastOnce AND xMixFound;
            END_IF

            o_stResult.xSuccess := o_xSuccess;

            (** 设置错误标志 **)
            IF xHasSingleError OR xHasMixError THEN
                o_xError := TRUE;
            END_IF

            (** 设置寻找结果标志 **)
            o_xSingleFound := xSingleFoundAtLeastOnce;
            o_xMixFound := xMixFound;

    END_CASE
END_IF

(** 设置报警标志 **)
o_xHasAlarm := xHasSingleError OR xHasMixError;
fbR_TRIG_HasAlarm(clk:=o_xHasAlarm);
IF fbR_TRIG_HasAlarm.Q THEN
	o_xHasAlarming:=TRUE;
END_IF
fbTON_HasAlarming(iN:=o_xHasAlarming,PT:=T#2000MS);
IF fbTON_HasAlarming.Q THEN
	fbTON_HasAlarming(iN:=FALSE);
	o_xHasAlarming:=FALSE;
END_IF

(** 更新全局数组 **)
FOR iN := 1 TO 3 BY 1 DO
	IF iN <= 2 THEN
		g_aiCurLabelPos[i_iAxisId, iN] := aiCurLabelPos[iN];
		g_arCurLabelWidth[i_iAxisId, iN] := arCurLabelWidth[iN];
		g_rFiberMoveDist[i_iAxisId, iN] := INT_TO_REAL((REAL_TO_INT(rFiberMoveDist[iN] * 10))) / 10;
	END_IF
	g_aiCurLabelPos[i_iAxisId, iN] := aiCurLabelPos[iN];
	g_arCurLabelWidth[i_iAxisId, iN] := arCurLabelWidth[iN];
END_FOR

g_aiStep_AutoAdjust[i_iAxisId] := eState;

o_stResult.eState:=eState;
(** 更新输出状态 **)
o_eState := eState;
o_xPressTriggered := xBeforeAxisPressTriggered;

(** 设置从站通信标志 **)
pstStRSV_UnitParam_UnSave^.byFlag_CommFromMaster.0 := i_xEn AND (eCmd <> FIND_CMD_RESET);
pstStRSV_UnitParam_UnSave^.byFlag_CommFromMaster.1 := o_xFindFirstMark;
pstStRSV_UnitParam_UnSave^.byFlag_CommFromMaster.3 := o_xFindPreMark;
pstStRSV_UnitParam_UnSave^.byFlag_CommFromMaster.5 := o_xGateMoveFinish;
pstStRSV_UnitParam_UnSave^.byFlag_CommFromMaster.6 := xMasterComplete;
pstStRSV_UnitParam_UnSave^.byFlag_CommFromMaster.7 := xFindMarkCenter_CalWidth;

(** 处理光纤移动 **)
pstStRSV_UnitParam_UnSave^.rFiberMoveDistanceIn_FindSignal := o_rFiberMoveDistanceIn_FindSignal;
pstStRSV_UnitParam_UnSave^.xFiberMoveDisRunStart_FindSignal := o_xFiberMoveDisRunStart_FindSignal;
IF ABS(o_rFiberMoveDistanceIn_FindSignal) < 0.1 THEN
    pstStRSV_UnitParam_UnSave^.xFiberMoveDisRunStart_FindSignal := FALSE;
END_IF
o_stResult.rFiberMoveDist:=o_rFiberMoveDistanceIn_FindSignal;
(*2026.05.21.095119上报金刚相关讯息||wang.xy*)
pstStRSV_UnitParam_UnSave^.wCommFromDubheFindSignal.0:=i_xEn AND (eCmd <> FIND_CMD_RESET);
pstStRSV_UnitParam_UnSave^.wCommFromDubheFindSignal.6 := xHasSingleError OR xHasMixError;
// pstStRSV_UnitParam_UnSave^.wCommFromDubheFindSignal.1:=
pstStRSV_UnitParam_UnSave^.iStep_AutoAdjust:=o_stResult.eState;
pstStRSV_UnitParam_UnSave^.iError_Msg:=o_stResult.iErrorCode;

// 					i_pstStSysParam^.astStRSV_UnitParam_UnSave[iUnitId].iStep_AutoAdjust;
// 	pstStParam_Diamonds_Wr_SysSts^.astStSts_UnitParam_2[iUnitId].iError_Msg:=
// 					i_pstStSysParam^.astStRSV_UnitParam_UnSave[iUnitId].iError_Msg;

(*日志*)
xNeedMsg :=FALSE;
IF eState<>ePrevState THEN
	tChangeStsTime:=TIME()-tLastTime;
	tLastTime:=TIME();
	//sTimeStamp_Tmp:= KS_GetTimeString(TIMEFORMAT_HYPHEN_DOT, TRUE, TRUE);
	sLogMsg := CONCAT('AXIS : ', INT_TO_STRING(i_iAxisId));
	sLogMsg := CONCAT(sLogMsg, '@');
	sLogMsg := CONCAT(sLogMsg, TIME_TO_STRING(tChangeStsTime));
	sLogMsg := CONCAT(sLogMsg,'|');
	sLogMsg := CONCAT(sLogMsg, INT_TO_STRING(ePrevState));
	sLogMsg := CONCAT(sLogMsg, '->');
	sLogMsg := CONCAT(sLogMsg, INT_TO_STRING(eState));
	xNeedMsg :=TRUE;
END_IF
(** 保存上一状态 **)
ePrevState := eState;

IF xNeedMsg THEN
	(* 调用日志函数 *)
	KS_HY_AddMsgToLog(
	g_pstStHYLogFifo,
	LOG_LEVEL_DEBUG,
	'MARKDETECTION',
	sLogMsg);
END_IF

(* ---- KS_FB_ManualFindMixColor.st ---- *)
(*@CES
Name=KS_FB_ManualFindMixColor
Type=FunctionBlock
TypeGuid=6f9dac99-8de1-4efc-8465-68ac443b7d08
Guid=48811e36-789b-45c0-9237-87d497c0d2dc
HasDeclaration=True
HasImplementation=True
*)
{DECLARATION}
FUNCTION_BLOCK KS_FB_ManualFindMixColor
VAR_INPUT
    i_iAxisId: INT;                      (* 轴号 *)
    i_pstStSysParam: POINTER TO StSysParam; (* 系统参数 *)
    i_rVel: REAL;                        (* 速度 *)
    i_rGirth: REAL;                      (* 版周长 *)
    i_rFilmLength: REAL;                 (* 料长 *)
    i_iBeforeAxisId: INT;                (* 前轴号（用于计算延时） *)
	i_pfbKS_FB_AxisFindModule: POINTER TO KS_FB_AxisFindModule;
END_VAR
VAR_OUTPUT
	o_xManualMixComplete :BOOL;           (*寻找完成*)
END_VAR
VAR
    pstStRSV_UnitParam_UnSave: POINTER TO StRSV_UnitParam_UnSave;
    pstStUnitParam_Save: POINTER TO StUnitParam_Save;
    pstStGrpParam_Save: POINTER TO StGrpParam_Save;
	pstStRSV_GrpParam_Save	: POINTER TO StRSV_GrpParam_Save;//
    rGirth: REAL;
    rFilmLength: REAL;
END_VAR

{IMPLEMENTATION}
(* 获取参数指针 *)
pstStRSV_UnitParam_UnSave := ADR(i_pstStSysParam^.astStRSV_UnitParam_UnSave[i_iAxisId]);
pstStUnitParam_Save := ADR(i_pstStSysParam^.astStUnitParam_Save[i_iAxisId]);
pstStGrpParam_Save:= ADR(i_pstStSysParam^.astStGrpParam_Save);
pstStRSV_GrpParam_Save :=  ADR(i_pstStSysParam^.astStRSV_GrpParam_Save);
rGirth := pstStUnitParam_Save^.rGirth_PrnRoller;
rFilmLength := pstStUnitParam_Save^.rFilmLengthFromPrevPressUnit;

(* 调用轴寻找模块 *)
i_pfbKS_FB_AxisFindModule^(
    (* 基本输入 *)
    i_xEn := TRUE,
    i_iAxisId := i_iAxisId,
    i_eCmd := FIND_CMD_START_MIX,
    i_xUseFindBestPosStep := FALSE,      (* 混色寻找不使用最佳位置步骤 *)

    (* 参数输入 *)
  	i_pstStRSV_UnitParam_UnSave := pstStRSV_UnitParam_UnSave,
	i_pstStUnitParam_Save := pstStUnitParam_Save,
	i_pstStGrpParam_Save := pstStGrpParam_Save,
    i_rVel := i_rVel,
    i_rGirth := rGirth,
    i_rFilmLength := rFilmLength,
    i_iBeforeAxisId := i_iBeforeAxisId,  (* 需要前轴号计算延时 *)
    i_iAfterAxisId := -1,                (* 手动模式不考虑后轴 *)
	i_rFindBestPos_MoveDis := pstStRSV_GrpParam_Save^.arFiberMove,

    (* 外部状态输入 *)
    i_xCoarseDone := TRUE,               (* 手动模式假设粗调已完成 *)
    i_xPressDone := TRUE,                (* 手动模式假设合压已完成 *)
    i_xAutoMode := FALSE,                (* 手动模式 *)
	i_xFind_IDLE := pstStRSV_UnitParam_UnSave^.byFlag_CommFromSlave.4,

    (* 开关参数 *)
    i_xSwitch_EnFastPress := FALSE,
    i_xSwitch_RFailure := FALSE,
    i_xSwitch_FFailure := FALSE,
    i_xSpecialMarkEn := FALSE
);

o_xManualMixComplete := i_pfbKS_FB_AxisFindModule^.o_xDone AND i_pfbKS_FB_AxisFindModule^.o_xSuccess;
